(* Logix 5000 project; controller DSFW_Budzar vendor 1 type 14 code 154 rev 32.13; software revision 32.03 *)
// Unit Model Number: DSFW-0512-C-FCB-S1-SP
// Unit Serial Number: 202008-38944-1

TASK MainTask (continuous, watchdog 500 ms) : A_MainProgram, B_Process_Control, D_Refrigeration_Control
TASK PID_Fast_Loop (periodic, rate 500 ms, priority 1, watchdog 1000 ms) : Pressure_PID, EEV_PID
TASK PID_Slow_Loop (periodic, rate 1000 ms, priority 1, watchdog 500 ms) : Main

MODULES
   Local : vendor 1 type 14 code 154 (PointIO 0, rev 32.13)
      SLOT_5 : 1734-IR2 (PointIO 5, rev 3.1, Input RPI 80 ms)
           Local:5:I.Ch0Data   // TE-105 Compressor Suction Temperature (404A)
           Local:5:I.Ch1Data   // TE-204 Evaporator Suction Line Temperature
      SLOT_4 : 1734-IR2 (PointIO 4, rev 3.1, Input RPI 80 ms)
           Local:4:I.Ch0Data   // TE-103 Liquid Line Temperature (404A)
           Local:4:I.Ch1Data   // TE-104 Evaporator Suction Temperature (404A)
      SLOT_2 : vendor 1 type 115 code 210 (PointIO 2, rev 3.1, Input RPI 80 ms)
           Local:2:I.Ch2Data   // PT-103 Compressor Discharge Pressure (449a)
           Local:2:I.Ch3Data   // PT-104 Evaporator Suction Line Pressure (449a)
           Local:2:I.Ch6Data   // PT-202 Evaporator Suction Line Pressure
           Local:2:I.Ch1Data   // PT-102 Compressor Suction Pressure (449a)
           Local:2:I.Ch0Data   // PT-101 Reactor Supply Pressure
           Local:2:I.Ch4Data   // PT-105 Nitrogen/Air Pressure
           Local:2:I.Ch7Data   // TT-*** Vessel Temperature
           Local:2:I.Ch5Data   // PT-201 Condenser Loop Supply Pressure
      SLOT_6 : 1734-IR2 (PointIO 6, rev 3.1, Input RPI 80 ms)
           Local:6:I.Ch0Data   // Spare
           Local:6:I.Ch1Data   // Spare
      SLOT_3 : 1734-IR2 (PointIO 3, rev 3.1, Input RPI 80 ms)
           Local:3:I.Ch0Data   // TE-101 Reactor Supply Temperature
           Local:3:I.Ch1Data   // TE-102 Reactor Return Temperature
      SLOT_9 : 1734-IE2C (PointIO 9, rev 3.1, Input RPI 80 ms)
           Local:9:I.Ch0Data   // FIT-101 Flow Indicating Transmitter
      Discrete_IO : Embedded (PointIO 1, rev 32.11, Output RPI 20 ms)
           Local:1:I.Data.0   // ESTOP
           Local:1:I.Data.1   // Phase Monitor
           Local:1:I.Data.10   // Spare
           Local:1:I.Data.11   // Spare
           Local:1:I.Data.12   // Compressor Low Oil Level
           Local:1:I.Data.13   // Condenser Loop Heater High Temperature Status
           Local:1:I.Data.14   // Condenser Loop Pump Run Proof Status
           Local:1:I.Data.15   // Spare
           Local:1:I.Data.2   // Purge Panel
           Local:1:I.Data.3   // Process Pump Run-Proof Contact
           Local:1:I.Data.4   // Process Heater #1 High Temperature
           Local:1:I.Data.5   // Spare
           Local:1:I.Data.6   // Spare
           Local:1:I.Data.7   // Spare
           Local:1:I.Data.8   // Compressor Run-Proof Contact
           Local:1:I.Data.9   // Compressor Motor Protector
           Local:1:O.Data.0   // Process Pump Motor Start Contactor
           Local:1:O.Data.1   // Process Heater #1 Output Enable
           Local:1:O.Data.10   // Spare
           Local:1:O.Data.11   // Spare
           Local:1:O.Data.12   // Spare
           Local:1:O.Data.13   // Spare
           Local:1:O.Data.14   // Spare
           Local:1:O.Data.15   // Spare
           Local:1:O.Data.2   // Spare
           Local:1:O.Data.3   // Spare
           Local:1:O.Data.4   // Spare
           Local:1:O.Data.5   // Compressor Motor Contactor
           Local:1:O.Data.6   // Spare
           Local:1:O.Data.7   // Spare
           Local:1:O.Data.8   // Condenser Loop Pump Motor Relay
           Local:1:O.Data.9   // Spare
      SLOT_8 : vendor 1 type 115 code 211 (PointIO 8, rev 3.1, Output RPI 80 ms)
           Local:8:O.Ch2Data   // Spare
           Local:8:O.Ch3Data   // Spare
           Local:8:O.Ch1Data   // PCV-101 Condenser Pressure Control
           Local:8:O.Ch0Data   // TCV-102 Hot Gas Bypass Valve
      SLOT_7 : vendor 1 type 115 code 211 (PointIO 7, rev 3.1, Output RPI 80 ms)
           Local:7:O.Ch2Data   // EEV-102 Compressor #1 Desuperheat Valve
           Local:7:O.Ch3Data   // TCV-101 Hot Gas Bypass Valve
           Local:7:O.Ch1Data   // EEV-101 Evaporator Electric Expansion Valve
           Local:7:O.Ch0Data   // SCR-101 SCR Heater Control
END_MODULES

TYPE BL_Analog_Input :
STRUCT
   Scale_4mA : REAL;
   Scale_20mA : REAL;
   Offset : REAL;
   Output : REAL;
   Fault_Delay : DINT;
END_STRUCT
END_TYPE

ADD_ON_INSTRUCTION BudLib_Analog_Sensor   (* revision 1.0 *)
VAR_IN_OUT
   BL_Analog_Input : BL_Analog_Input; {required}
END_VAR
VAR_INPUT
   Raw_Data : REAL; {required}
   Sensor_Type : BOOL; {required}   // 0 = 4-20mA 1 = RTD
   Disable_High_Fault : BOOL; {required}
END_VAR
VAR_OUTPUT
   Sensor_Alarm : BOOL; {access None, required}
END_VAR
VAR_INPUT
   CLR_Alarm : BOOL; {required}
   Fault_Disable : BOOL; {required}   // Disable Fault
END_VAR
VAR
   Fault_Delay_TMR : TIMER; {access None}
END_VAR

ROUTINE Logic   (* ladder *)
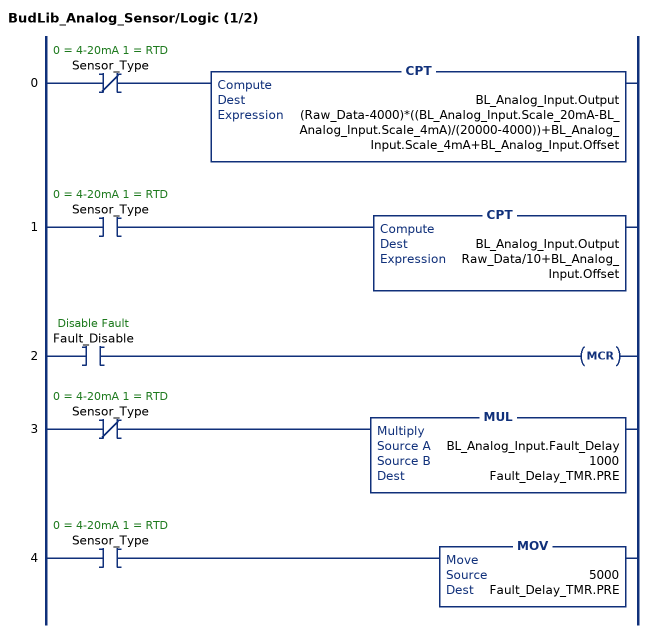
   0: XIO(Sensor_Type)CPT(BL_Analog_Input.Output,(Raw_Data-4000)*((BL_Analog_Input.Scale_20mA-BL_Analog_Input.Scale_4mA)/(20000-4000))+BL_Analog_Input.Scale_4mA+BL_Analog_Input.Offset);
   1: XIC(Sensor_Type)CPT(BL_Analog_Input.Output,Raw_Data/10+BL_Analog_Input.Offset);
   2: XIC(Fault_Disable)MCR();
   3: XIO(Sensor_Type)MUL(BL_Analog_Input.Fault_Delay,1000,Fault_Delay_TMR.PRE);
   4: XIC(Sensor_Type)MOV(5000,Fault_Delay_TMR.PRE);
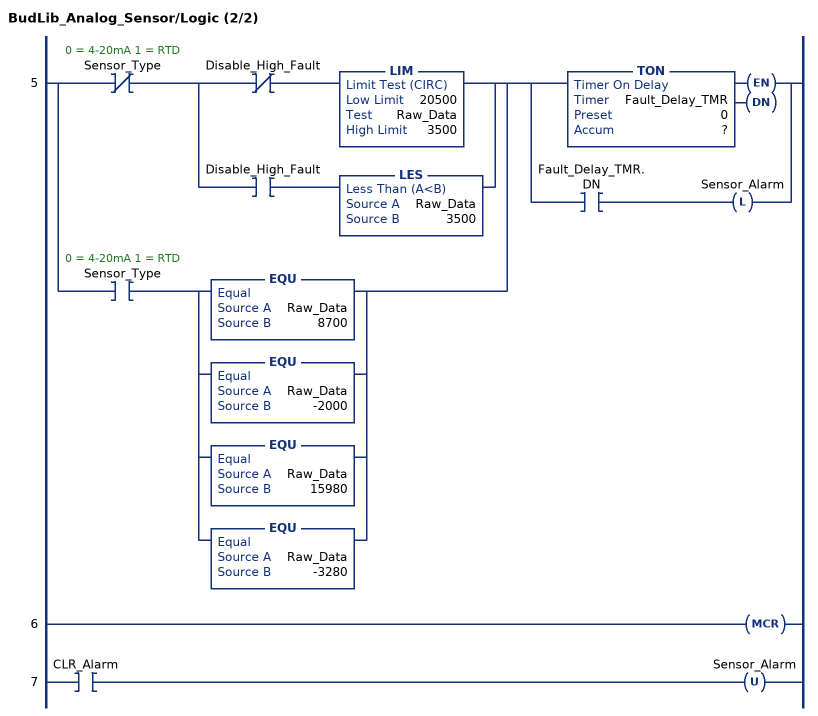
   5: [XIO(Sensor_Type) [XIO(Disable_High_Fault) LIM(20500,Raw_Data,3500) ,XIC(Disable_High_Fault) LES(Raw_Data,3500) ] ,XIC(Sensor_Type) [EQU(Raw_Data,8700) ,EQU(Raw_Data,-2000) ,EQU(Raw_Data,15980) ,EQU(Raw_Data,-3280) ] ][TON(Fault_Delay_TMR,?,?) ,XIC(Fault_Delay_TMR.DN) OTL(Sensor_Alarm) ];
   6: MCR();
   7: XIC(CLR_Alarm)OTU(Sensor_Alarm);
END_ROUTINE
END_ADD_ON_INSTRUCTION

ADD_ON_INSTRUCTION BudLib_Compressor   (* revision 1.0 *)
// Compressor Cycle and Antirecycle
VAR_OUTPUT
   PLC_Address : BOOL; {access Read Only, required}   // Compressor Start Relay
END_VAR
VAR_INPUT
   Start_Delay_Time : DINT; {required}   // Minimum Off Time, (milliseconds)
   Short_Cycle_Time : DINT; {required}   // Short Cycle Time (milliseconds)
END_VAR
VAR_OUTPUT
   Time_Remaining : DINT; {access Read Only, required}
   Compressor_Timing : BOOL; {access Read Only, required}
END_VAR
VAR_INPUT
   Compressor_OK_TO_RUN : BOOL; {access Read Only, required}
END_VAR
VAR_OUTPUT
   Start_Delay_DN : BOOL; {access Read Only}
   Start_Delay_EN : BOOL; {access Read Only}
   Start_Delay_Remaining : DINT; {access Read Only}
END_VAR
VAR
   Short_Cycle_TMR : TIMER; {access None}   // Short Cycle Timer
   Start_TMR : TIMER; {access None}   // Start Delay Timer
END_VAR

ROUTINE Logic   (* ladder *)
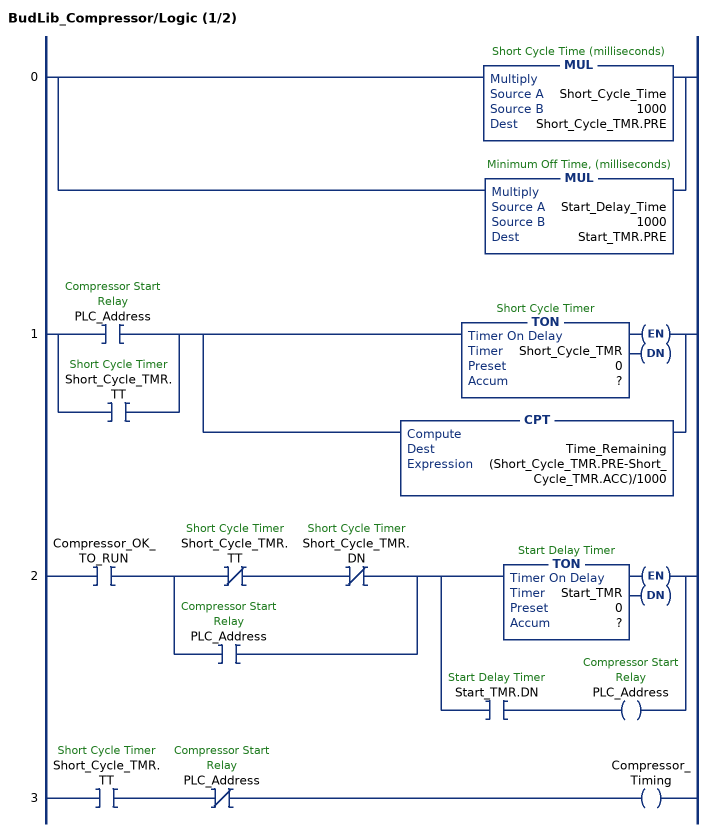
   0: [MUL(Short_Cycle_Time,1000,Short_Cycle_TMR.PRE) ,MUL(Start_Delay_Time,1000,Start_TMR.PRE) ];
   1: [XIC(PLC_Address) ,XIC(Short_Cycle_TMR.TT) ][TON(Short_Cycle_TMR,?,?) ,CPT(Time_Remaining,(Short_Cycle_TMR.PRE-Short_Cycle_TMR.ACC)/1000) ];
   2: XIC(Compressor_OK_TO_RUN)[XIO(Short_Cycle_TMR.TT) XIO(Short_Cycle_TMR.DN) ,XIC(PLC_Address) ][TON(Start_TMR,?,?) ,XIC(Start_TMR.DN) OTE(PLC_Address) ];
   3: XIC(Short_Cycle_TMR.TT)XIO(PLC_Address)OTE(Compressor_Timing);
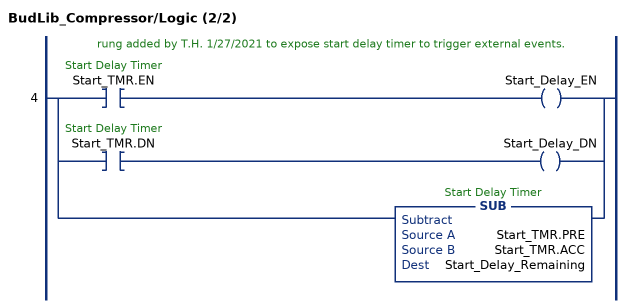
   // rung added by T.H. 1/27/2021 to expose start delay timer to trigger external events.
   4: [XIC(Start_TMR.EN) OTE(Start_Delay_EN) ,XIC(Start_TMR.DN) OTE(Start_Delay_DN) ,SUB(Start_TMR.PRE,Start_TMR.ACC,Start_Delay_Remaining) ];
END_ROUTINE
END_ADD_ON_INSTRUCTION

ADD_ON_INSTRUCTION BudLib_Heater_Step_Controller   (* revision 1.0, vendor Budzar Industries, Inc. *)
// Heaters Step Controller For Up To 10 Heaters
// Revision note:
// Initial Release 20Dec2017 (cdz)
VAR_IN_OUT
   Power_Request : REAL; {required}   // Heaters Power Request From TIC
   Heater_Circuits : DINT; {required}   // Number Of Heaters To Control (Includes SCR Controlled Heater)
   SCR : DINT; {required}   // Output To SCR scaled 0% to 100% Power
   Heater_Contactors : DINT; {required}   // Heater Contactors ON Commands (Interlock Individual Heater Circuits Outside AOI)
END_VAR
VAR_INPUT
   Interlock : BOOL; {required}   // Instruction Interlock (Sets All Outputs To Zero)
END_VAR
VAR
   Power_Total : DINT; {access None}   // Internal Calculation
   Step_Power : DINT[11]; {access None}   // Internal Calculation
END_VAR

ROUTINE Logic   (* ladder *)
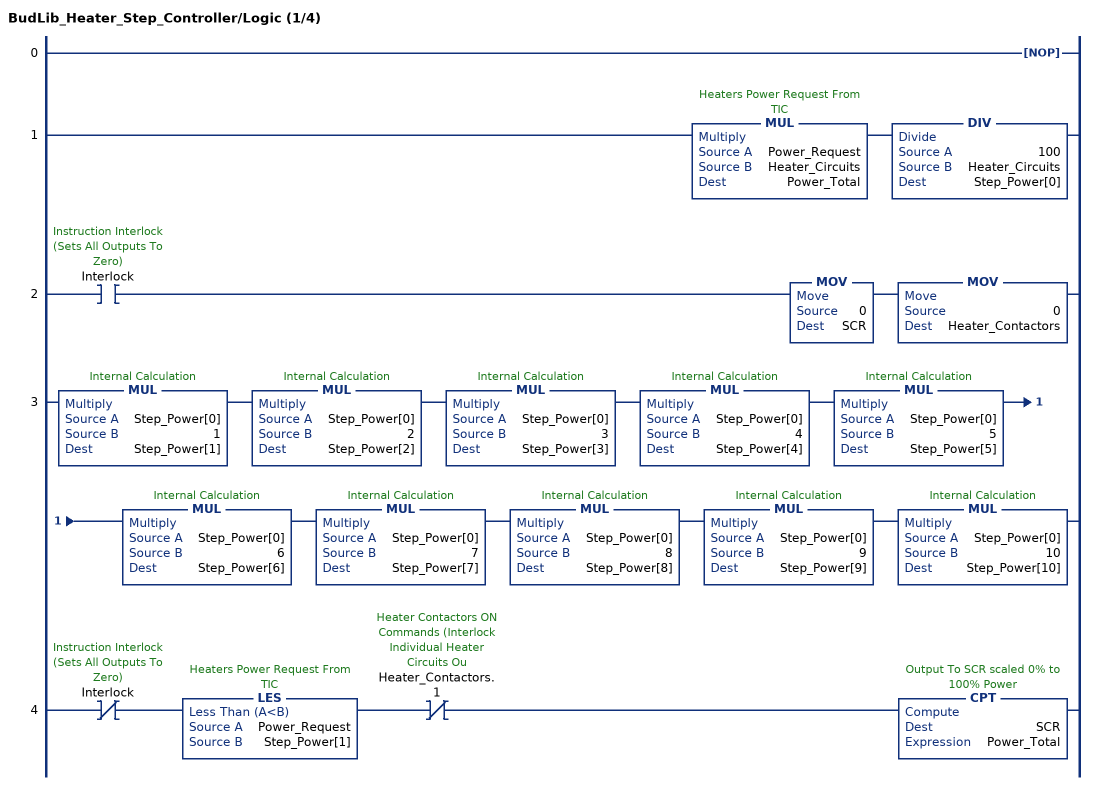
   0: NOP();
   1: MUL(Power_Request,Heater_Circuits,Power_Total)DIV(100,Heater_Circuits,Step_Power[0]);
   2: XIC(Interlock)MOV(0,SCR)MOV(0,Heater_Contactors);
   3: MUL(Step_Power[0],1,Step_Power[1])MUL(Step_Power[0],2,Step_Power[2])MUL(Step_Power[0],3,Step_Power[3])MUL(Step_Power[0],4,Step_Power[4])MUL(Step_Power[0],5,Step_Power[5])MUL(Step_Power[0],6,Step_Power[6])MUL(Step_Power[0],7,Step_Power[7])MUL(Step_Power[0],8,Step_Power[8])MUL(Step_Power[0],9,Step_Power[9])MUL(Step_Power[0],10,Step_Power[10]);
   4: XIO(Interlock)LES(Power_Request,Step_Power[1])XIO(Heater_Contactors.1)CPT(SCR,Power_Total);
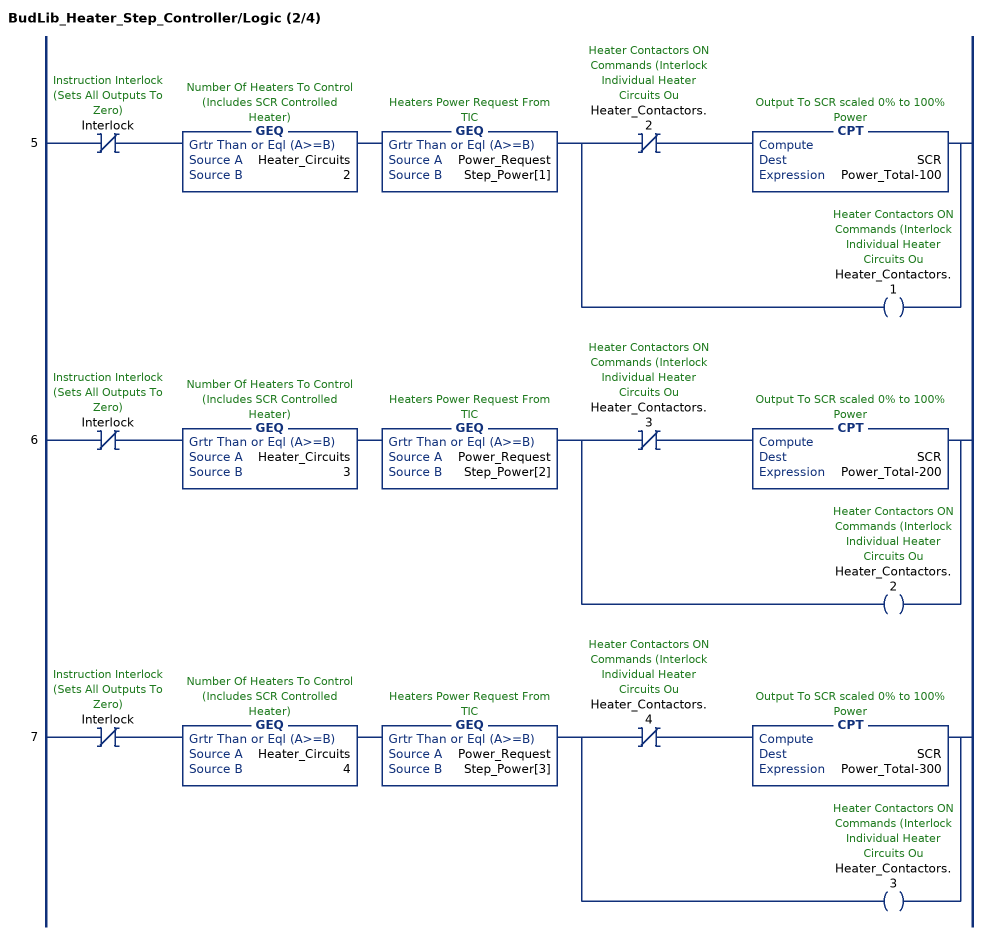
   5: XIO(Interlock)GEQ(Heater_Circuits,2)GEQ(Power_Request,Step_Power[1])[XIO(Heater_Contactors.2) CPT(SCR,Power_Total-100) ,OTE(Heater_Contactors.1) ];
   6: XIO(Interlock)GEQ(Heater_Circuits,3)GEQ(Power_Request,Step_Power[2])[XIO(Heater_Contactors.3) CPT(SCR,Power_Total-200) ,OTE(Heater_Contactors.2) ];
   7: XIO(Interlock)GEQ(Heater_Circuits,4)GEQ(Power_Request,Step_Power[3])[XIO(Heater_Contactors.4) CPT(SCR,Power_Total-300) ,OTE(Heater_Contactors.3) ];
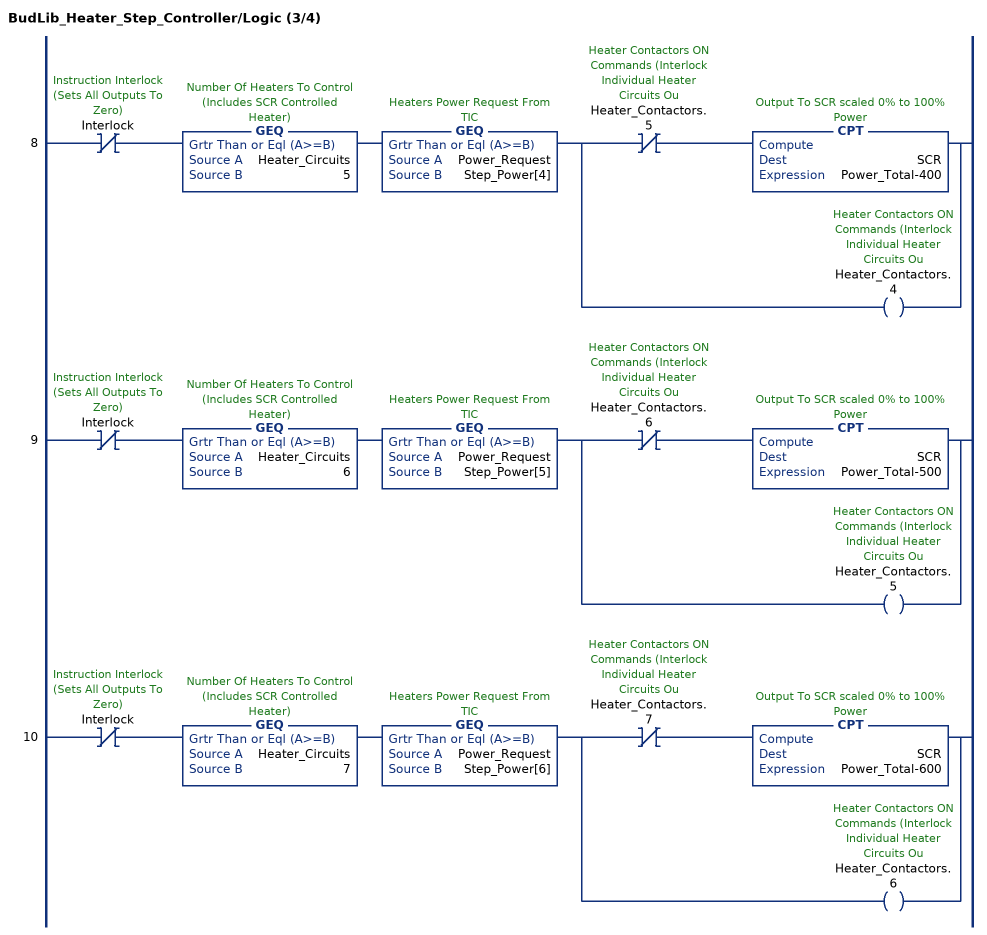
   8: XIO(Interlock)GEQ(Heater_Circuits,5)GEQ(Power_Request,Step_Power[4])[XIO(Heater_Contactors.5) CPT(SCR,Power_Total-400) ,OTE(Heater_Contactors.4) ];
   9: XIO(Interlock)GEQ(Heater_Circuits,6)GEQ(Power_Request,Step_Power[5])[XIO(Heater_Contactors.6) CPT(SCR,Power_Total-500) ,OTE(Heater_Contactors.5) ];
   10: XIO(Interlock)GEQ(Heater_Circuits,7)GEQ(Power_Request,Step_Power[6])[XIO(Heater_Contactors.7) CPT(SCR,Power_Total-600) ,OTE(Heater_Contactors.6) ];
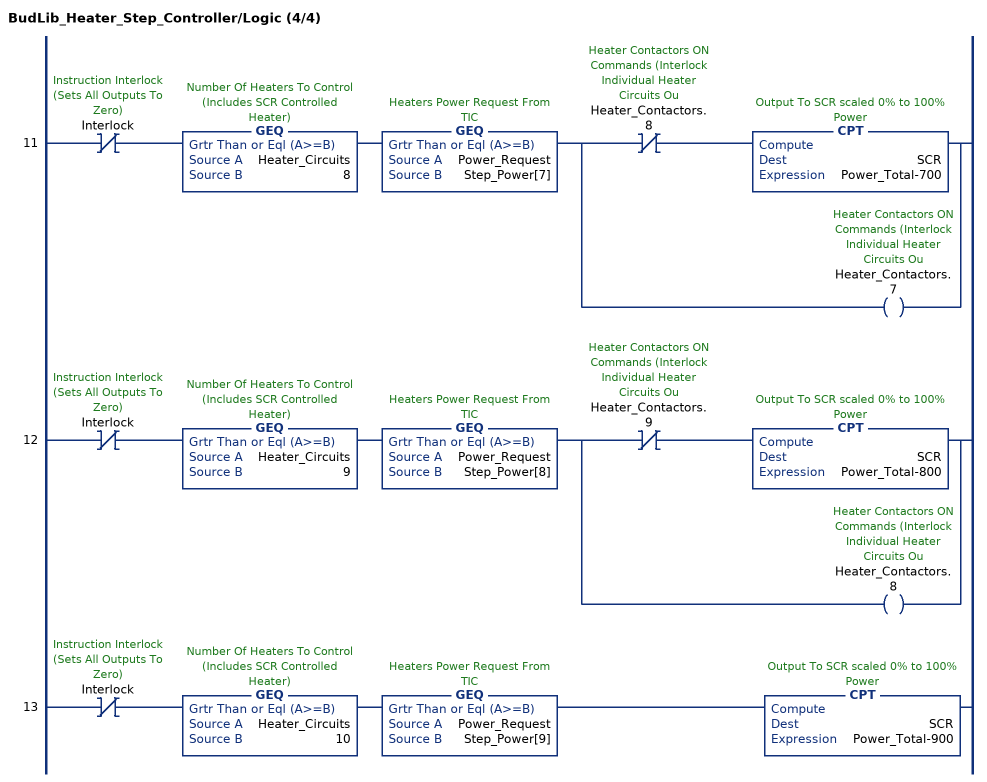
   11: XIO(Interlock)GEQ(Heater_Circuits,8)GEQ(Power_Request,Step_Power[7])[XIO(Heater_Contactors.8) CPT(SCR,Power_Total-700) ,OTE(Heater_Contactors.7) ];
   12: XIO(Interlock)GEQ(Heater_Circuits,9)GEQ(Power_Request,Step_Power[8])[XIO(Heater_Contactors.9) CPT(SCR,Power_Total-800) ,OTE(Heater_Contactors.8) ];
   13: XIO(Interlock)GEQ(Heater_Circuits,10)GEQ(Power_Request,Step_Power[9])CPT(SCR,Power_Total-900);
END_ROUTINE
END_ADD_ON_INSTRUCTION

ADD_ON_INSTRUCTION BudLib_Superheat_Subcooling   (* revision 1.2 *)
// Revision note:
// Added Refrigerant 508B
// Added Refrigerant R449A
VAR_INPUT
   Temperature : REAL; {required}   // Suction or Liquid Line Temperature
   Pressure : REAL; {required}   // Suction or Discharge Pressure
END_VAR
VAR_OUTPUT
   P2T_Suction : REAL; {access Read Only}   // Suction Pressure to Temperature Calculation
   P2T_Liquid : REAL; {access Read Only}   // Liquid Pressure to Temperature Calculation
END_VAR
VAR_INPUT
   Refridgerant_Type : INT; {required}   // 1=R-22 2=R-134a 3=R-404a 4=R-407c 5=R-407a 6=R-410a 7=R-422d 8=R-438a 9=R-507 10=R-508B 11=R-449A 12=R290
   Superheat_Subcool : BOOL; {required}   // 0 = Superheat, 1 = Subcool
END_VAR
VAR_OUTPUT
   Result : REAL; {required}   // Calculated Result
END_VAR
VAR
   Superheat : REAL; {access Read Only}   // Superheat Calculation
   Subcool : REAL; {access Read Only}   // Subcool Calculation
END_VAR

ROUTINE Logic   (* structured text *)
   
   
   Case Refridgerant_Type OF
   
   (* R-22 *)
   1:  P2T_Suction:= -0.000000165*Pressure**4 + 0.000084606*Pressure**3 - 0.016568240*Pressure**2 + 1.952262699*Pressure - 39.085397206;
       P2T_Liquid:= -0.000000165*Pressure**4 + 0.000084606*Pressure**3 - 0.016568240*Pressure**2 + 1.952262699*Pressure - 39.085397206;
   
   (*R-134a*)
   2: P2T_Suction:= -0.00000000000037678795*Pressure**6 + 0.00000000056931121499*Pressure**5 - 0.00000033878300479892*Pressure**4 + 0.00010202087796451500*Pressure**3 - 0.01710716970609380000*Pressure**2 + 1.97485706462976000*Pressure - 12.16021651744090;
      P2T_Liquid:= -0.00000000000037678795*Pressure**6 + 0.00000000056931121499*Pressure**5 - 0.00000033878300479892*Pressure**4 + 0.00010202087796451500*Pressure**3 - 0.01710716970609380000*Pressure**2 + 1.97485706462976000*Pressure - 12.16021651744090;
   
   (*R-404a*)
   3:  P2T_Suction:= -0.00000000005300893321*Pressure**6 + 0.00000002741449672112*Pressure**5 - 0.00000570303468006017*Pressure**4 + 0.00062421870492102000*Pressure**3 - 0.04148675026965520000*Pressure**2 + 2.37637660990731000000*Pressure - 49.68565233808480000000;
       P2T_Liquid:= -0.0000000000000550315164227*Pressure**6 + 0.0000000000997514242404528*Pressure**5 - 0.0000000737248710163770000*Pressure**4 + 0.0000290410699131178000000*Pressure**3- 0.0069198966935964100000000*Pressure**2  + 1.2825072984089100*Pressure - 33.916124534865200;
   
   (*R-407c*)
   4:   P2T_Suction := -0.00000000000800924737*Pressure**6 + 0.00000000557131285962*Pressure**5 - 0.00000169384905437941*Pressure**4 + 0.00028593017513500700*Pressure**3 - 0.02893370732670060000*Pressure**2 + 2.20060661934258000000*Pressure - 33.32183919094680000000;
   	P2T_Liquid:= 0.00000000000002386292*Pressure**6 - 0.00000000002645317402*Pressure**5 + 0.00000000526050718724*Pressure**4 + 0.00000470562626432580*Pressure**3 - 0.00310591635937629000*Pressure**2 + 1.00142167143801000000*Pressure - 22.25895791216770000000;
   
   (*R-407a*)
   5:	P2T_Suction:= -0.00000000011518362850*Pressure**6 + 0.00000005009100701803*Pressure**5 - 0.00000875403007261077*Pressure**4 + 0.00080807995686882400*Pressure**3 - 0.04608857801110840000*Pressure**2 + 2.36986927227190000000*Pressure - 37.26735163389090000000;
   	P2T_Liquid:= -0.00000000000003784489*Pressure**6 + 0.00000000006834533715*Pressure**5 - 0.00000005140162309636*Pressure**4 + 0.00002127640311370790*Pressure**3 - 0.00554724395898896000*Pressure**2 + 1.16486749118176000000*Pressure - 30.11932356915960000000;
   
   (*R-410a*)
   6:	P2T_Suction:= -0.00000000000007186775*Pressure**6 + 0.00000000014583668666*Pressure**5 - 0.00000011674472220023*Pressure**4 + 0.00004726707063285040*Pressure**3 - 0.01057489539488190000*Pressure**2 + 1.57409368233857000000*Pressure - 56.17353301327970000000;
   	P2T_Liquid:= -0.00000000000007186775*Pressure**6 + 0.00000000014583668666*Pressure**5 - 0.00000011674472220023*Pressure**4 + 0.00004726707063285040*Pressure**3 - 0.01057489539488190000*Pressure**2 + 1.57409368233857000000*Pressure - 56.17353301327970000000;
   
   (*R-422D*)
   7:	P2T_Suction:= 0.00000000056957976185*Pressure**5 - 0.00000058362559681170*Pressure**4 + 0.00016582335662478100*Pressure**3 - 0.02207715168838590000*Pressure**2 + 2.02610656700961000000*Pressure - 35.18819939281650000000;
   	P2T_Liquid:= 0.00000000000813454044*Pressure**5 - 0.00000001433073228086*Pressure**4 + 0.00001015786430530350*Pressure**3 - 0.00389055376093068000*Pressure**2 + 1.06625906617128000000*Pressure - 22.58790116749710000000;
   
   (*R-438a*)
   8:	P2T_Suction:= 0.00000000006078715896*Pressure**6 - 0.00000001611318229885*Pressure**5 + 0.00000020938844025320*Pressure**4 + 0.00027696642267471800*Pressure**3 - 0.03274545521389880000*Pressure**2 + 2.29322301382490000000*Pressure - 32.72178606997110000000;
   	P2T_Liquid:=  -0.00000000000003163289*Pressure**6 + 0.00000000006045751232*Pressure**5 - 0.00000004802369289111*Pressure**4 + 0.00002089758452796680*Pressure**3 - 0.00566402177639559000*Pressure**2 + 1.20642331219452000000*Pressure - 25.80440294280620000000;
   
   (*R-507*)
   9:	P2T_Suction:= -0.00000000000023273589*Pressure**6 + 0.00000000038440242299*Pressure**5 - 0.00000024966416650859*Pressure**4 + 0.00008180023458648210*Pressure**3 - 0.01483731477723890000*Pressure**2 + 1.83216631968571000000*Pressure - 49.09858575703400000000;
   	P2T_Liquid:=  -0.00000000000023273589*Pressure**6 + 0.00000000038440242299*Pressure**5 - 0.00000024966416650859*Pressure**4 + 0.00008180023458648210*Pressure**3 - 0.01483731477723890000*Pressure**2 + 1.83216631968571000000*Pressure - 49.09858575703400000000;
   
   (*R-508B*)
   10:	P2T_Suction:= -0.000000000000133667762*Pressure**6 + 0.000000000236822589*Pressure**5 - 0.000000165498946*Pressure**4 + 0.0000585053021*Pressure**3 - 0.01144174*Pressure**2 + 1.5057373*Pressure - 123.74624;
   	P2T_Liquid:=  -0.000000000000133667762*Pressure**6 + 0.000000000236822589*Pressure**5 - 0.000000165498946*Pressure**4 + 0.0000585053021*Pressure**3 - 0.01144174*Pressure**2 + 1.5057373*Pressure - 123.74624;
   
   (*R-449A*)
   11: P2T_Suction:= -0.00000000000036541159*Pressure**6 + 0.00000000054907825576*Pressure**5 - 0.00000032708993709514*Pressure**4 + 0.00009916804470212850*Pressure**3 - 0.01675694050709890000*Pressure**2 + 1.91534370751567000000*Pressure - 39.0570030049292;
   	P2T_Liquid:=  -0.00000000000036907278*Pressure**6 + 0.00000000055456970769*Pressure**5 - 0.00000033032085879095*Pressure**4 + 0.00010012437901080800*Pressure**3 - 0.01690317434666350000*Pressure**2 + 1.93545495275924000000*Pressure - 49.96916448983160000000;
   
   (*R-290*)
   12: P2T_Suction:= -8.90208426e-013*Pressure**6 + 1.11806286e-009*Pressure**5 - 5.57465512e-007*Pressure**4 + 1.42291974e-004*Pressure**3 - 0.020612964*Pressure**2 + 2.1470945*Pressure - 41.50468;
       P2T_Liquid := -8.90208426e-013*Pressure**6 + 1.11806286e-009*Pressure**5 - 5.57465512e-007*Pressure**4 + 1.42291974e-004*Pressure**3 - 0.020612964*Pressure**2 + 2.1470945*Pressure - 41.50468;
   
   END_CASE;
   
   
   IF NOT Superheat_Subcool THEN
   	Superheat:=Temperature - P2T_Suction;
   	Result := Superheat;
   
   ELSE
   	Subcool:= P2T_Liquid - Temperature;
   	Result := Subcool;
   
   END_IF;
END_ROUTINE
END_ADD_ON_INSTRUCTION

ADD_ON_INSTRUCTION P2T   (* revision 1.1 *)
// Revision note:
// Added Refrigerant 508B
VAR_INPUT
   SuctionRTD : REAL; {required}   // Suction Line RTD
   LiquidRTD : REAL; {required}   // Liquid Line RTD
   Suction_Pressure : REAL; {required}   // Compressor Suction Pressure
   Discharge_Pressure : REAL; {required}   // Compressor Discharge Pressure
END_VAR
VAR_OUTPUT
   P2T_Suction : REAL; {access Read Only}   // Suction Pressure to Temperature Calculation
   Superheat : REAL; {access Read Only, required}   // Superheat Calculation
   P2T_Liquid : REAL; {access Read Only}   // Liquid Pressure to Temperature Calculation
   Subcool : REAL; {access Read Only, required}   // Subcool Calculation
END_VAR
VAR_INPUT
   Refridgerant_Type : INT; {required}   // 1=R-22 2=R-134a 3=R-404a 4=R-407c 5=R-407a 6=R-410a 7=R-422d 8=R-438a 9=R-507 10=R-508B
END_VAR

ROUTINE Logic   (* structured text *)
   
   
   Case Refridgerant_Type OF
   
   (* R-22 *)
   1:  P2T_Suction:= -0.000000165*Suction_Pressure**4 + 0.000084606*Suction_Pressure**3 - 0.016568240*Suction_Pressure**2 + 1.952262699*Suction_Pressure - 39.085397206;
       P2T_Liquid:= -0.000000165*Discharge_Pressure**4 + 0.000084606*Discharge_Pressure**3 - 0.016568240*Discharge_Pressure**2 + 1.952262699*Discharge_Pressure - 39.085397206; ;
   
   (*R-134a*)
   2: P2T_Suction:= -0.00000000000037678795*Suction_Pressure**6 + 0.00000000056931121499*Suction_Pressure**5 - 0.00000033878300479892*Suction_Pressure**4 + 0.00010202087796451500*Suction_Pressure**3 - 0.01710716970609380000*Suction_Pressure**2 + 1.97485706462976000*Suction_Pressure - 12.16021651744090;
      P2T_Liquid:= -0.00000000000037678795*Discharge_Pressure**6 + 0.00000000056931121499*Discharge_Pressure**5 - 0.00000033878300479892*Discharge_Pressure**4 + 0.00010202087796451500*Discharge_Pressure**3 - 0.01710716970609380000*Discharge_Pressure**2 + 1.97485706462976000*Discharge_Pressure - 12.16021651744090;
   
   (*R-404a*)
   3:  P2T_Suction:= -0.00000000005300893321*Suction_Pressure**6 + 0.00000002741449672112*Suction_Pressure**5 - 0.00000570303468006017*Suction_Pressure**4 + 0.00062421870492102000*Suction_Pressure**3 - 0.04148675026965520000*Suction_Pressure**2 + 2.37637660990731000000*Suction_Pressure - 49.68565233808480000000;
       P2T_Liquid:= -0.0000000000000550315164227*Discharge_Pressure**6 + 0.0000000000997514242404528*Discharge_Pressure**5 - 0.0000000737248710163770000*Discharge_Pressure**4 + 0.0000290410699131178000000*Discharge_Pressure**3- 0.0069198966935964100000000*Discharge_Pressure**2  + 1.2825072984089100*Discharge_Pressure - 33.916124534865200;
   
   (*R-407c*)
   4:   P2T_Suction := -0.00000000000800924737*Suction_Pressure**6 + 0.00000000557131285962*Suction_Pressure**5 - 0.00000169384905437941*Suction_Pressure**4 + 0.00028593017513500700*Suction_Pressure**3 - 0.02893370732670060000*Suction_Pressure**2 + 2.20060661934258000000*Suction_Pressure - 33.32183919094680000000;
   	P2T_Liquid:= 0.00000000000002386292*Discharge_Pressure**6 - 0.00000000002645317402*Discharge_Pressure**5 + 0.00000000526050718724*Discharge_Pressure**4 + 0.00000470562626432580*Discharge_Pressure**3 - 0.00310591635937629000*Discharge_Pressure**2 + 1.00142167143801000000*Discharge_Pressure - 22.25895791216770000000;
   
   (*R-407a*)
   5:	P2T_Suction:= -0.00000000011518362850*Suction_Pressure**6 + 0.00000005009100701803*Suction_Pressure**5 - 0.00000875403007261077*Suction_Pressure**4 + 0.00080807995686882400*Suction_Pressure**3 - 0.04608857801110840000*Suction_Pressure**2 + 2.36986927227190000000*Suction_Pressure - 37.26735163389090000000;
   	P2T_Liquid:= -0.00000000000003784489*Discharge_Pressure**6 + 0.00000000006834533715*Discharge_Pressure**5 - 0.00000005140162309636*Discharge_Pressure**4 + 0.00002127640311370790*Discharge_Pressure**3 - 0.00554724395898896000*Discharge_Pressure**2 + 1.16486749118176000000*Discharge_Pressure - 30.11932356915960000000;
   
   (*R-410a*)
   6:	P2T_Suction:= -0.00000000000007186775*Suction_Pressure**6 + 0.00000000014583668666*Suction_Pressure**5 - 0.00000011674472220023*Suction_Pressure**4 + 0.00004726707063285040*Suction_Pressure**3 - 0.01057489539488190000*Suction_Pressure**2 + 1.57409368233857000000*Suction_Pressure - 56.17353301327970000000;
   	P2T_Liquid:= -0.00000000000007186775*Discharge_Pressure**6 + 0.00000000014583668666*Discharge_Pressure**5 - 0.00000011674472220023*Discharge_Pressure**4 + 0.00004726707063285040*Discharge_Pressure**3 - 0.01057489539488190000*Discharge_Pressure**2 + 1.57409368233857000000*Discharge_Pressure - 56.17353301327970000000;
   
   (*R-422D*)
   7:	P2T_Suction:= 0.00000000056957976185*Suction_Pressure**5 - 0.00000058362559681170*Suction_Pressure**4 + 0.00016582335662478100*Suction_Pressure**3 - 0.02207715168838590000*Suction_Pressure**2 + 2.02610656700961000000*Suction_Pressure - 35.18819939281650000000;
   	P2T_Liquid:= 0.00000000000813454044*Discharge_Pressure**5 - 0.00000001433073228086*Discharge_Pressure**4 + 0.00001015786430530350*Discharge_Pressure**3 - 0.00389055376093068000*Discharge_Pressure**2 + 1.06625906617128000000*Discharge_Pressure - 22.58790116749710000000;
   
   (*R-438a*)
   8:	P2T_Suction:= 0.00000000006078715896*Suction_Pressure**6 - 0.00000001611318229885*Suction_Pressure**5 + 0.00000020938844025320*Suction_Pressure**4 + 0.00027696642267471800*Suction_Pressure**3 - 0.03274545521389880000*Suction_Pressure**2 + 2.29322301382490000000*Suction_Pressure - 32.72178606997110000000;
   	P2T_Liquid:=  -0.00000000000003163289*Discharge_Pressure**6 + 0.00000000006045751232*Discharge_Pressure**5 - 0.00000004802369289111*Discharge_Pressure**4 + 0.00002089758452796680*Discharge_Pressure**3 - 0.00566402177639559000*Discharge_Pressure**2 + 1.20642331219452000000*Discharge_Pressure - 25.80440294280620000000;
   
   (*R-507*)
   9:	P2T_Suction:= -0.00000000000023273589*Suction_Pressure**6 + 0.00000000038440242299*Suction_Pressure**5 - 0.00000024966416650859*Suction_Pressure**4 + 0.00008180023458648210*Suction_Pressure**3 - 0.01483731477723890000*Suction_Pressure**2 + 1.83216631968571000000*Suction_Pressure - 49.09858575703400000000;
   	P2T_Liquid:=  -0.00000000000023273589*Discharge_Pressure**6 + 0.00000000038440242299*Discharge_Pressure**5 - 0.00000024966416650859*Discharge_Pressure**4 + 0.00008180023458648210*Discharge_Pressure**3 - 0.01483731477723890000*Discharge_Pressure**2 + 1.83216631968571000000*Discharge_Pressure - 49.09858575703400000000;
   
   (*R-508B*)
   10:	P2T_Suction:= -0.000000000000133667762*Suction_Pressure**6 + 0.000000000236822589*Suction_Pressure**5 - 0.000000165498946*Suction_Pressure**4 + 0.0000585053021*Suction_Pressure**3 - 0.01144174*Suction_Pressure**2 + 1.5057373*Suction_Pressure - 123.74624;
   	P2T_Liquid:=  -0.000000000000133667762*Discharge_Pressure**6 + 0.000000000236822589*Discharge_Pressure**5 - 0.000000165498946*Discharge_Pressure**4 + 0.0000585053021*Discharge_Pressure**3 - 0.01144174*Discharge_Pressure**2 + 1.5057373*Discharge_Pressure - 123.74624;
   
   
   END_CASE;
   
   Superheat:=SuctionRTD - P2T_Suction;
   
   Subcool:= P2T_Liquid - LiquidRTD;
   
END_ROUTINE
END_ADD_ON_INSTRUCTION

VAR_GLOBAL   (* controller tags *)
   ACKNOWLEDGE_ALARMS : BOOL;
   Active_Setpoint : REAL := 20.0;
   ALARMS : DINT[5] := ([1] := 2#0000_0001_0000_0000_0000_0000_0000_0000);
        [0]   // SENSOR ALARMS
        [0].0   // PT-101 Process Supply Pressure Sensor Fault
        [0].1   // PT-102 404A Compressor Suction Pressure Sensor Fault
        [0].10   // TE-101 Process Supply Temperature Sensor Fault
        [0].11   // TE-102 Process Return Temperature Sensor Fault
        [0].12   // TE-103 404A Liquid Line Temperature Sensor Fault
        [0].13   // TE-104 404A Evaporator Suction Temperature Sensor Fault
        [0].14   // TE-105 404A Compressor Suction Temperature Sensor Fault
        [0].15   // TE-106 Condenser Chilled Water Outlet Temperature Sensor Fault
        [0].16   // TE-108 Condenser Chilled Water Inlet Temperature Sensor Fault
        [0].2   // PT-103 404A Compressor Discharge Pressure Sensor Fault
        [0].3   // PT-104 404A Evaporator Suction Line Pressure Sensor Fault
        [0].4   // PT-105 4 MTR-101 Low Suction Pressure Sensor Fault
        [0].5   // FIT-101 Process Supply Flow Transmitter Fault
        [0].6   // PT-107 Pump Suction Pressure Sensor Fault
        [0].7   // PT-108 Pump Discharge Pressure Sensor Fault
        [0].9   // TT-*** Vessel Temperature Transmitter Sensor Fault
        [1]   // General/Process Alarms
        [1].0   // Process Pump Run-Proof Alarm
        [1].1   // Heater #1 Elements High Temperature Alarm
        [1].10   // Jacket High High Temperature Alarm
        [1].11   // Jacket HighTemperature Alarm
        [1].12   // Vessel Low Low Temperature Alarm
        [1].13   // Spare
        [1].14   // Vessel High High Temperature Alarm
        [1].15   // Jacket/Vessel High Delta T Alarm
        [1].16   // Glycol Tank Low Level Alarm
        [1].17   // Process Pump Low Suction Pressure Alarm
        [1].18   // Spare
        [1].19   // Spare
        [1].2   // Spare
        [1].20   // Purge Panel Low Pressure
        [1].21   // Spare
        [1].23   // Remote Temperature Setpoint from Plant DCS is out-of-range
        [1].24   // DCS Communication Fault
        [1].25   // Condenser Water Inlet Temperature High Alarm
        [1].3   // Phase Monitor Fault
        [1].4   // Emergency Stop
        [1].5   // Process Pump Low Pressure Alarm
        [1].6   // Process Pump High Pressure Alarm
        [1].8   // Jacket Low Low Temperature Alarm
        [1].9   // Jacket Low Temperature Alarm
        [2]   // R404A Refrigeration Alarms
        [2].0   // Compressor Run-Proof Alarm
        [2].1   // Compressor Low Pressure
        [2].11   // PT-202 CONDENSER EVAPORATOR SUCTION LINE PRESSURE TRANSMITTER ALARM
        [2].12   // TE-201 CONDENSER LOOP SUPPLY TEMPERATURE SENSOR FAULT
        [2].13   // TE-202 CONDENSER LOOP RETURN TEMPERATURE SENSOR FAULT
        [2].14   // TE-204 EVAPORATOR SUCTION LINE TEMPERATURE SENSOR FAULT
        [2].2   // Compressor High Pressure
        [2].3   // Low Superheat
        [2].4   // High Superheat
        [2].5   // Compressor Low Oil Level
        [2].6   // Compressor Motor Protector
        [2].7   // Condening Glycol/Water Temmperature Too High Alarm
        [4]   // Module Faults
        [4].0   // PLC101 SLOT 2 1734-IE8C MODULE CRASH
        [4].1   // PLC101 SLOT 3 1734-IR2 MODULE CRASH
        [4].2   // PLC101 SLOT 4 1734-IR2 MODULE CRASH
        [4].3   // PLC101 SLOT 5 1734-IR2 MODULE CRASH
        [4].4   // PLC101 SLOT 6 1734-IR2 MODULE CRASH
        [4].5   // PLC101 SLOT 7 1734-OE4C MODULE CRASH
        [4].6   // PLC101 SLOT 8 1734-OE4C MODULE CRASH
        [4].7   // PLC101 SLOT 9 1734-IE2C MODULE CRASH
   ALARMS_PRESENT : BOOL := 1;
   ALWAYS_OFF : BOOL;
   Batch_High_High_Temp_Delay : TIMER := (PRE := 30000);
   Batch_High_High_Temp_Setpoint : REAL;
   Batch_High_Temp_Setpoint : REAL;
   Batch_Jacket_DT_Temp_Delay : TIMER := (PRE := 30000);
   Batch_Low_Low_Temp_Delay : TIMER := (PRE := 30000);
   Batch_Low_Low_Temp_Setpoint : REAL := -10.0;
   Batch_Low_Temp_Delay : TIMER := (PRE := 5000);
   Batch_Low_Temp_Setpoint : REAL;
   Batch_Mode_Enable : BOOL;
   Batch_Mode_Running : BOOL;
   Blanket_Pressure_Delta_PV : REAL := 0.95624924;
   BudLib_P2T_1 : BudLib_Superheat_Subcooling := (Temperature := 85.1, Pressure := 110.7004, P2T_Suction := 53.529312, P2T_Liquid := 53.13972, Refridgerant_Type := 3, Result := 31.570686);
   BudLib_P2T_2 : BudLib_Superheat_Subcooling := (Temperature := 73.7, Pressure := 163.45125, P2T_Suction := 73.087265, P2T_Liquid := 75.620316, Refridgerant_Type := 3, Superheat_Subcool := 1, Result := 1.9203186);
   BudLib_P2T_3 : BudLib_Superheat_Subcooling := (Temperature := 75.1, Pressure := 110.693596, P2T_Suction := 53.524734, P2T_Liquid := 53.136364, Refridgerant_Type := 3, Result := 21.575264);
   BudLib_P2T_4 : BudLib_Superheat_Subcooling := (Temperature := 26.4, Pressure := 24.42431, P2T_Suction := -9.100571, P2T_Liquid := -6.3220596, Refridgerant_Type := 3, Result := 35.500572);
   C1_Low_Oil_Timer : TIMER := (PRE := 5000);
   C1_MP_Timer : TIMER := (PRE := 3000);
   C1_Run_Proof_Timer : TIMER := (PRE := 3000);
   C2_MP_Timer : TIMER := (PRE := 3000);
   C2_Run_Proof_Timer : TIMER := (PRE := 3000);
   C3_MP_Timer : TIMER := (PRE := 3000);
   C3_Run_Proof_Timer : TIMER := (PRE := 3000);
   C_101_AUX : ALIAS FOR Local:1:I.Data.8;
   CLR_Alarms : BOOL;
   Comp_1 : BudLib_Compressor := (Start_Delay_Time := 10, Short_Cycle_Time := 300, Start_Delay_Remaining := 10000);   // R507A Compressor 1
   Comp_1_Status : BOOL;
   Comp_404A_Timing_1 : BOOL;
   Comp_404A_Timing_2 : BOOL;
   Comp_Start_Purge_Relay : BOOL;
   Compressor_R404A_Subcooling : REAL := 1.9203186;
   Compressor_R404A_Superheat : REAL := 31.570686;
   Compressor_Start_Request : BOOL;
   Condenser_Water_Inlet_Temp_Limit : REAL := 100.0;
   Condenser_Water_Inlet_Temp_TMR : TIMER := (PRE := 10000);
   CR_002 : ALIAS FOR Local:1:I.Data.0;   // Emergency Stop Safety Relay Status
   CR_003 : ALIAS FOR Local:1:O.Data.15;   // General Fault Relay
   CR_01 : ALIAS FOR Local:1:I.Data.15;   // Glycol Tank Low Level Alarm Relay Dry Contact
   CR_108 : ALIAS FOR Local:1:O.Data.0;   // Process Pump Motor Relay (Energizes Contactor M-101)
   CR_109 : ALIAS FOR Local:1:O.Data.5;   // Compressor Motor Relay (Energizes Contactor C-101)
   CR_201 : ALIAS FOR Local:1:O.Data.8;   // GFS-10 Auto Start Relay (Enables Glycol Pump)
   DCS_Comm_TMR : TIMER := (PRE := 10000, ACC := 10000, EN := 1, DN := 1);
   DCS_Heartbeat_Returned : DINT;
   DCS_Heartbeat_Returned_Last : DINT;
   EEV_101_Auto_Manual : BOOL;
   EEV_101_High_Range_CV_Max : REAL := 65.0;
   EEV_101_High_Range_CV_Min : REAL := 9.0;
   EEV_101_Low_Range_CV_Max : REAL := 88.0;
   EEV_101_Low_Range_CV_Min : REAL := 5.0;
   EEV_101_Manual_Percent : REAL := 100.0;
   EEV_101_Mid_Range_CV_Max : REAL := 87.0;
   EEV_101_Mid_Range_CV_Min : REAL := 8.0;
   EEV_101_Pressure_PIDE : PID_ENHANCED := (PV := 110.693596, PVEUMax := 121.5, PVEUMin := -27.3, SPProg := 100.0, SPOper := 100.0, SPHLimit := 121.5, SPLLimit := -27.3, RatioProg := 1.0, RatioOper := 1.0, RatioHLimit := 1.0, RatioLLimit := 1.0, CVEUMax := 20000.0, CVEUMin := 4000.0, CVHLimit := 87.0, CVLLimit := 8.0, HandFB := 100.0, PGain := 3.0, IGain := 8.0, PVEDerivative := 1, ProgOverrideReq := 1, RTSTime := 1, CVEU := 4000.0, CVLAlarm := 1, SP := 100.0, SPPercent := 85.55108, PVPercent := 92.737625, E := -10.693596, EPercent := -7.1865463, InitPrimary := 1, WindupLOut := 1, Ratio := 1.0, ProgOper := 1, Override := 1, DeltaT := 0.5);
   EEV_101_Pressure_Setpoint : REAL := 100.0;
   EEV_101_Run_PIDE : BOOL;
   EEV_101_Run_Temp_PIDE : BOOL;
   EEV_101_SH_PIDE : PID_ENHANCED := (PV := 21.575264, PVEUMax := 200.0, PVEUMin := -100.0, SPProg := 12.0, SPOper := 12.0, SPHLimit := 200.0, SPLLimit := -100.0, RatioProg := 1.0, RatioOper := 1.0, RatioHLimit := 1.0, RatioLLimit := 1.0, CVEUMax := 20000.0, CVEUMin := 4000.0, CVHLimit := 87.0, CVLLimit := 8.0, HandFB := 100.0, ControlAction := 1, PGain := 5.0, IGain := 12.0, PVEDerivative := 1, ProgOverrideReq := 1, RTSTime := 1, CVEU := 4000.0, CVLAlarm := 1, SP := 12.0, SPPercent := 37.333332, PVPercent := 40.52509, E := 9.575264, EPercent := 3.1917572, InitPrimary := 1, WindupHOut := 1, Ratio := 1.0, ProgOper := 1, Override := 1, DeltaT := 0.5);
   EEV_101_Stop_PIDE : BOOL := 1;
   EEV_101_Superheat_Setpoint : REAL := 12.0;
   EEV_101_Temperature_PIDE : PID_ENHANCED := (PV := 23.3, PVEUMax := 200.0, PVEUMin := -40.0, SPProg := 20.0, SPOper := 23.3, SPCascade := 23.3, SPHLimit := 200.0, SPLLimit := -40.0, RatioProg := 1.0, RatioOper := 1.0, RatioHLimit := 1.0, RatioLLimit := 1.0, CVEUMax := 20000.0, CVEUMin := 4000.0, CVHLimit := 87.0, CVLLimit := 8.0, HandFB := 100.0, ControlAction := 1, PGain := 3.0, IGain := 8.0, PVEDerivative := 1, PVTracking := 1, AllowCasRat := 1, ProgOverrideReq := 1, RTSTime := 1, CVEU := 4000.0, CVLAlarm := 1, SP := 23.3, SPPercent := 26.374998, PVPercent := 26.374998, InitPrimary := 1, WindupHOut := 1, Ratio := 1.0, ProgOper := 1, Override := 1, DeltaT := 0.5);
   EEV_101_To_Purge : BOOL;   // Oil Management, Call For Purge with EEV-101
   EEV_102_Auto_Manual : BOOL;
   EEV_102_Manual_Percent : REAL;
   EEV_102_PIDE : PID_ENHANCED := (PV := 31.570686, PVEUMax := 200.0, PVEUMin := -40.0, SPProg := 40.0, SPOper := 31.570686, SPHLimit := 200.0, SPLLimit := -40.0, RatioProg := 1.0, RatioOper := 1.0, RatioHLimit := 1.0, RatioLLimit := 1.0, CVEUMax := 20000.0, CVEUMin := 4000.0, CVHLimit := 100.0, ControlAction := 1, PGain := 2.0, IGain := 3.0, PVEDerivative := 1, PVTracking := 1, ProgOverrideReq := 1, RTSTime := 1, CVEU := 4000.0, SP := 31.570686, SPPercent := 29.82112, PVPercent := 29.82112, InitPrimary := 1, Ratio := 1.0, ProgOper := 1, Override := 1, DeltaT := 0.5);
   EEV_102_Run_PIDE : BOOL;
   EEV_102_Stop_PIDE : BOOL := 1;
   EEV_102_Superheat_Setpoint : REAL := 40.0;
   EEV_201_Auto_Manual : BOOL;
   EEV_High_Range_Max_Temp : REAL := 90.0;
   EEV_High_Range_Min_Temp : REAL := 55.1;
   EEV_Low_Range_Max_Temp : REAL := -5.0;
   EEV_Low_Range_Min_Temp : REAL := -10.0;
   EEV_Manual_Relief_Delay : TIMER := (PRE := 75000);   // Oil Management, Delay until Flush begins
   EEV_Manual_Relief_Timer : TIMER := (PRE := 15000);   // Oil Management, Duration of Flush
   EEV_Mid_Range_Max_Temp : REAL := 55.0;
   EEV_Mid_Range_Min_Temp : REAL := -4.1;
   Enable_Batch : BOOL;   // Batch/Jacket Mode 0=Jacket 1=Batch
   Engineering_Alarm_Reset : TIMER := (PRE := 10000);
   Evaporator_R404A_Superheat : REAL := 21.575264;
   F8 : REAL[48] := ([0] := 24.885624, [2] := 0.033749998, [3] := 22.1, [5] := 23.3, [6] := 25.1575, [7] := 24.813124, [8] := 110.693596, [9] := 75.1, [10] := 85.1, [11] := 110.7004, [12] := 73.7, [13] := 163.45125, [14] := 73.4, [15] := 28.827812, [16] := 71.5, [17] := 47.85, [23] := 20.0, [28] := 25.0); {produced}   // FLOAT DATA FOR PLANT SUPERVISORY SYSTEM
   FCV_101 : ALIAS FOR Local:8:O.Ch2Data;   // Process Bypass Flow Control Valve
   FIC_101_Manual_Percent : REAL := 50.0;
   FIC_101_PIDE : PID_ENHANCED := (PV := 0.031875, PVEUMax := 165.0, PVEUMin := -20.0, SPProg := 20.0, SPOper := 0.031875, SPHLimit := 165.0, SPLLimit := -20.0, RatioProg := 1.0, RatioOper := 1.0, RatioHLimit := 1.0, RatioLLimit := 1.0, CVEUMax := 20000.0, CVEUMin := 4000.0, CVHLimit := 100.0, HandFB := 50.0, PGain := 1.2, IGain := 25.0, PVEDerivative := 1, PVTracking := 1, ProgOverrideReq := 1, RTSTime := 1, CVEU := 4000.0, SP := 0.031875, SPPercent := 10.82804, PVPercent := 10.82804, InitPrimary := 1, Ratio := 1.0, ProgOper := 1, Override := 1, DeltaT := 0.5);
   FIC_101_Run_PID : BOOL;
   FIC_101_Setpoint : REAL := 20.0;
   FIC_101_Stop_PID : BOOL := 1;
   FIT_101 : BL_Analog_Input := (Scale_20mA := 30.0, Output := 0.031875);   // Flow Indicating Transmitter
   FIT_101_PID_Scale_Max : REAL := 165.0;
   FIT_101_PID_Scale_Min : REAL := -20.0;
   Glycol_Pump_Disable_TMR : TIMER := (PRE := 10000);   // Disable Glycol Fill Pump on High PSI (backup for Pressure Switch on Neptune)
   Heater_Contactors : DINT;
   Heater_Step_Controller : BudLib_Heater_Step_Controller := (Interlock := 1);
   High_Range_Max_Temp : REAL := 90.0;
   High_Range_Min_Temp : REAL := 55.1;
   HMI_Batch_Hi_Hi_Temp_Delay : DINT := 30;
   HMI_Batch_Jacket_DT_Temp_Delay : DINT := 30;
   HMI_Batch_Low_Low_Temp_Delay : DINT := 30;
   HMI_Bypass_Speed : DINT := 3;
   HMI_Bypass_Status : BOOL;
   HMI_Condenser_Water_Inlet_Temp_Delay : DINT := 10;
   HMI_EEV_101_CV : REAL;
   HMI_EEV_101_Lamp : BOOL;
   HMI_EEV_102_CV : REAL;
   HMI_EEV_102_Lamp : BOOL;
   HMI_EEV_Manual_Relief_Delay : REAL := 75.0;   // Oil Management, Delay to start relief entered in minutes.
   HMI_EEV_Manual_Relief_Timer : REAL := 15.0;   // Oil Management, Relief Duration entered in seconds
   HMI_FCV_101_CV : REAL;
   HMI_FCV_101_Lamp : BOOL;
   HMI_Heater_1_Lamp : BOOL;
   HMI_Heater_2_Lamp : BOOL;
   HMI_Jacket_Hi_Hi_Temp_Delay : DINT := 30;
   HMI_Jacket_Hi_Temp_Delay : REAL := 30.0;
   HMI_Jacket_Low_Low_Temp_Delay : DINT := 30;
   HMI_Jacket_Low_Temp_Delay : REAL := 30.0;
   HMI_Low_Pump_Suction_Pressure_Delay : REAL := 30.0;
   HMI_Low_Suction_Pressure_Delay : DINT := 10;
   HMI_Oil_Purge_Retries_Reset_Min : REAL := 10.0;   // Oil Management, Compressor Runtime before resetting retry accumulator
   HMI_PCV_101_Flush_Time : DINT := 30;
   HMI_PCV_101_Lamp : BOOL;
   HMI_PCV_101_Output : REAL;
   HMI_Pump_Start : BOOL;
   HMI_Pump_Status : BOOL;
   HMI_Pump_Stop : BOOL;
   HMI_R404A_Hot_Gas_Switch_Delay : REAL := 10.0;
   HMI_R404A_TCV_Toggle_SP : REAL := 60.0;
   HMI_R404A_Valve_Flush_SP : REAL := 80.0;   // Oil Management, desired valve position for Flush (0-100%)
   HMI_R507A_High_Superheat_Timer : DINT := 120;
   HMI_R507A_Low_Pressure_Delay : DINT := 120;
   HMI_R507A_Low_Superheat_Timer : DINT := 120;
   HMI_Ramping : BOOL;
   HMI_Remote_State_1 : BOOL;
   HMI_Remote_State_2 : BOOL;
   HMI_Return_Trend_Limits : REAL[2] := ([0] := -7.8999996, [1] := 52.1);
   HMI_SCR_Max : DINT;
   HMI_Soaking : BOOL;
   HMI_SP_Trend_Limits : REAL[2] := ([0] := -10.0, [1] := 50.0);
   HMI_Supply_Flow_Speed : DINT := 3;
   HMI_Supply_Flow_Status : BOOL;
   HMI_Supply_Trend_Limits : REAL[2] := ([0] := -6.700001, [1] := 53.3);
   HMI_TCV_101_CV : REAL;
   HMI_TCV_101_Lamp : BOOL;
   HMI_TCV_102_CV : REAL;
   HMI_TCV_102_Lamp : BOOL;
   HMI_TCV_Manual_Relief_Delay : REAL := 60.0;
   HMI_TCV_Manual_Relief_Timer : REAL := 10.0;
   HMI_Trend_Data : REAL[3] := ([0] := 20.0, [1] := 23.3, [2] := 22.1);
        [0]   // Temperature Setpoint
        [1]   // Process Supply Temperature
        [2]   // Process Return Temperature
   HMI_Valve_Flush_SP : REAL := 60.0;
   Jacket_Batch_Delta_T : REAL := 132.44063;
   Jacket_Batch_High_Delta_T_Setpoint : REAL := 100.0;
   Jacket_High_High_Temp_Delay : TIMER := (PRE := 30000);
   Jacket_High_High_Temp_Setpoint : REAL := 100.0;
   Jacket_High_Temp_Delay : TIMER := (PRE := 30000);
   Jacket_High_Temp_Setpoint : REAL := 90.0;
   Jacket_Low_Low_Temp_Delay : TIMER := (PRE := 30000);
   Jacket_Low_Low_Temp_Setpoint : REAL := -20.0;
   Jacket_Low_Temp_Delay : TIMER := (PRE := 30000);
   Jacket_Low_Temp_Setpoint : REAL := -10.0;
   Local_System_Start : BOOL;   // Local System Start 0=Stop 1=Start
   Local_Temp_Setpoint : REAL := 20.0;   // Local Temperature Setpoint
   Low_Pump_Suction_Pressure_Delay : TIMER := (PRE := 30000);
   Low_Pump_Suction_Pressure_Setpoint : REAL := 4.0;
   Low_Range_Max_Temp : REAL;
   Low_Range_Min_Temp : REAL := -10.0;
   M_101_AUX : ALIAS FOR Local:1:I.Data.3;
   Mid_Range_Max_Temp : REAL := 55.0;
   Mid_Range_Min_Temp : REAL := 0.1;
   N7 : INT[16] := ([0] := 26, [1] := 32, [10] := 60, [11] := 2); {produced}   // INTEGER DATA FOR PLANT SUPERVISORY SYSTEM
        [11].0   // REMOTE START PUSH BUTTON
        [11].1   // REMOTE STOP PUSH BUTTON
   New_Alarm_TMR : TIMER := (PRE := 500);
   NEW_ALARMS : DINT[5];   // New Alarms this scan
   NEW_ALARMS_PRESENT : BOOL;   // New Alarm Present This Scan
   NOT_ALARMS_LAST : DINT[5] := ([0] := -1, [1] := -16777217, [2] := -1, [3] := -1, [4] := -1);   // Logical NOT of Alarms Last Scan
   Num_Heaters : DINT := 2;
   Oil_Purge_Fail : BOOL;   // Oil Management, This coil will energize after configured purge retries fail
   Oil_Purge_Relay : BOOL;   // Oil Management, Oil Purge Sequence Latch
   Oil_Purge_Retires_Enable : BOOL;
   Oil_Purge_Retries_ACC : DINT;   // Oil Management, Accumulated Oil Purges this low level
   Oil_Purge_Retries_Reset : TIMER := (PRE := 600000);   // Oil Management, Reset Accumulator with 10-min without Low Level
   Oil_Purge_Retries_Reset1 : TIMER := (PRE := 10000, ACC := 10002, EN := 1, DN := 1);   // Oil Management, Used to reset accuulated retries if compressor off.
   Oil_Purge_Retries_Reset_Remaining : REAL;   // Oil Management, Time remaining until reset retries accum
   Oil_Purge_Retries_SP : DINT := 6;   // Oil Management, Desired Oil Purge Retries before Fault
   OMB_101 : ALIAS FOR Local:1:I.Data.12;
   ONS : DINT[3] := ([0] := 5);   // One-Shots
   P2T_507A : P2T := (SuctionRTD := 66.4, LiquidRTD := 61.8, Suction_Pressure := 76.8296, Discharge_Pressure := 124.46438, P2T_Suction := 34.86673, Superheat := 31.533272, P2T_Liquid := 59.58862, Subcool := -2.21138, Refridgerant_Type := 3);
   PCV_101_Auto_Manual : BOOL;
   PCV_101_Condenser_Pressure_PIDE : PID_ENHANCED := (PV := 163.45125, PVEUMax := 455.0, PVEUMin := -20.0, SPProg := 150.0, SPOper := 163.45125, SPHLimit := 455.0, SPLLimit := -20.0, RatioProg := 1.0, RatioOper := 1.0, RatioHLimit := 1.0, RatioLLimit := 1.0, CVEUMax := 20000.0, CVEUMin := 4000.0, CVHLimit := 100.0, HandFB := 100.0, ControlAction := 1, PGain := 4.0, IGain := 40.0, PVEDerivative := 1, PVTracking := 1, ProgOverrideReq := 1, RTSTime := 1, CVEU := 4000.0, SP := 163.45125, SPPercent := 38.621315, PVPercent := 38.621315, InitPrimary := 1, Ratio := 1.0, ProgOper := 1, Override := 1, DeltaT := 0.5);
   PCV_101_Flush_Limit : REAL := 70.0;   // Temperature Limit (Deg F) to force Condenser Water Flush
   PCV_101_Flush_Position : REAL := 20000.0;   // PCV-101 Desired Flush Position (4000-20000 counts)
   PCV_101_Flush_Time_Remaining : DINT := 30;
   PCV_101_Flush_Timer : TIMER := (PRE := 30000);   // PCV-101 Condenser Hot Water Flush Timer
   PCV_101_go_to_start_position : BOOL;
   PCV_101_Manual_Output : REAL := 100.0;
   PCV_101_Multiplexer : DINT := 1;   // Selects controlling input to multiplxer
   PCV_101_Pressure_SP : REAL := 150.0;
   PCV_101_Run_PIDE : BOOL;
   PCV_101_Start_Position : REAL := 12000.0;   // PCV-101 Desired Start Position (4000-20000 counts)
   PCV_101_Stop_PIDE : BOOL := 1;
   PLC_DateTime : DINT[7] := ([0] := 2026, [1] := 8, [2] := 24, [3] := 17, [4] := 17, [5] := 26, [6] := 851406);
        [0]   // year
        [1]   // month
        [2]   // day
        [3]   // hour
        [4]   // minute
        [5]   // seconds
        [6]   // microseconds
   PM_101 : ALIAS FOR Local:1:I.Data.1;
   PM_101_StartupTMR : TIMER := (PRE := 30000, ACC := 30002, EN := 1, DN := 1);   // PM-101 Phase Monitor Startup Delay Alarm Timer
   Process_Pump_Diff_Pressure : REAL := -3.960312;
   PT_101 : BL_Analog_Input := (Scale_20mA := 145.0, Output := 24.930937, Fault_Delay := 5);   // Process Supply Pressure
   PT_102 : BL_Analog_Input := (Scale_4mA := -7.3, Scale_20mA := 101.5, Output := 110.7004);   // R404A Compressor Suction Pressure
   PT_102_PID_Scale_Max : REAL := 121.5;
   PT_102_PID_Scale_Min : REAL := -27.3;
   PT_103 : BL_Analog_Input := (Scale_20mA := 435.0, Output := 163.45125, Fault_Delay := 5);   // R404A Compressor Discharge Pressure
   PT_103_PID_Scale_Max : REAL := 455.0;
   PT_103_PID_Scale_Min : REAL := -20.0;
   PT_104 : BL_Analog_Input := (Scale_4mA := -7.3, Scale_20mA := 101.5, Output := 110.693596);   // R404A Evaporator Suction Pressure
   PT_104_PID_Scale_Max : REAL := 121.5;
   PT_104_PID_Scale_Min : REAL := -27.3;
   PT_105 : BL_Analog_Input := (Scale_20mA := 145.0, Output := 28.855);   // Condenser Chilled Glycol Return Pressure
   PT_106 : BL_Analog_Input := (Scale_20mA := 145.0, Output := 47.868122);   // Condenser Chilled Glycol Supply Pressure
   PT_107 : BL_Analog_Input := (Scale_20mA := 145.0, Output := 25.1575);   // Process Pump Suction Pressure
   PT_108 : BL_Analog_Input := (Scale_20mA := 145.0, Output := 24.813124);   // Process Pump Suction Discharge Pressure
   Pump_1_Low_Press_Delay : TIMER := (PRE := 30000);
   Pump_High_Pressure_Alarm_Setpoint : REAL := 120.0;
   Pump_Low_Pressure_Alarm_Setpoint : REAL := 10.0;
   Pump_Manual_Release : BOOL := 1;
   Pump_Manual_Release_Timer : TIMER := (PRE := 5000, ACC := 5001, EN := 1, DN := 1);
   Pump_OK_To_Run : BOOL := 1;
   Pump_RP_ALM_TMR : TIMER := (PRE := 3000);
   Pump_Running : BOOL;
   Purge_Request : BOOL;   // Oil Management, Request to Purge
   R404A_HG_Switch_Delay : TIMER := (PRE := 10000);
   R404A_HG_Switch_Off_Delay : TIMER := (PRE := 10000);
   R404A_High_Pressure_Setpoint : REAL := 350.0;
   R404A_High_SH_Setpoint : REAL := 80.0;
   R404A_High_Superheat_Timer : TIMER := (PRE := 120000);
   R404A_Hot_Gas_Toggle : BOOL;
   R404A_Hot_Gas_Toggle_Req : BOOL;
   R404A_Low_Pressure_Delay : TIMER := (PRE := 120000);
   R404A_Low_Pressure_Setpoint : REAL := 15.0;
   R404A_Low_SC_Setpoint : REAL;
   R404A_Low_SH_Setpoint : REAL := 2.0;
   R404A_Low_Subcooling_Timer : TIMER := (PRE := 120000);
   R404A_Low_Superheat_Timer : TIMER := (PRE := 120000);
   R404A_Oil_Purge_Retires_Enable : BOOL;   // Oil Management, Oil Purge Retries Enabled
   R404A_OK_To_Run : BOOL;
   R404A_One_Comp_Running : BOOL;
   R404A_TCV_Toggle_SP_OFF : REAL := 58.0;
   R404A_TCV_Toggle_SP_ON : REAL := 62.0;
   R404A_TCV_Valve_Toggle : BOOL;
   Ramp_Soak_Current_HMI : DINT := 2#0000_0000_0000_0000_0000_0000_0000_0001;
   Ramp_Soak_Segments_HMI : DINT := 2#0000_0000_0000_0000_0000_0000_0011_1110;
   Ramp_Soak_Segments_HMI_Set : REAL := 5.0;
   REACTOR_BATCH_PID_START : BOOL;
   REACTOR_BATCH_PID_STOP : BOOL := 1;
   REACTOR_BATCH_PIDE : PID_ENHANCED := (PV := 20.0, PVEUMax := 200.0, PVEUMin := -40.0, SPProg := 20.0, SPOper := 20.0, SPHLimit := 200.0, SPLLimit := -40.0, RatioProg := 1.0, RatioOper := 1.0, RatioHLimit := 1.0, RatioLLimit := 1.0, CVInitReq := 1, CVInitValue := 23.3, CVOper := 51.454544, CVEUMax := 50.0, CVEUMin := -5.0, CVHLimit := 100.0, PGain := 12.0, IGain := 4.0, PVEDerivative := 1, DSmoothing := 1, PVTracking := 1, AllowCasRat := 1, ProgOverrideReq := 1, RTSTime := 1, CVEU := 23.3, CV := 51.454544, CVInitializing := 1, SP := 20.0, SPPercent := 25.0, PVPercent := 25.0, InitPrimary := 1, Ratio := 1.0, Override := 1, DeltaT := 1.0);
   REACTOR_BATCH_PIDE_CV_AS_SP : REAL := 23.3;
   REACTOR_BATCH_PV : REAL := 20.0;
   REACTOR_BATCH_SP_HIGH : REAL := 50.0;
   REACTOR_BATCH_SP_LOW : REAL := -10.0;
   REACTOR_HEAT_RUN_PIDE : BOOL;
   REACTOR_HEAT_STOP_PIDE : BOOL := 1;
   REACTOR_HEATERS_OK_TO_RUN : BOOL;
   REACTOR_HEATERS_TEMPERATURE_PIDE : PID_ENHANCED := (PV := 23.3, PVEUMax := 200.0, PVEUMin := -40.0, SPProg := 20.0, SPOper := 23.3, SPCascade := 23.3, SPHLimit := 200.0, SPLLimit := -40.0, RatioProg := 1.0, RatioOper := 1.0, RatioHLimit := 1.0, RatioLLimit := 1.0, CVEUMax := 20000.0, CVEUMin := 4000.0, CVHLimit := 100.0, HandFB := 78.0, PGain := 12.0, IGain := 3.0, PVEDerivative := 1, PVTracking := 1, AllowCasRat := 1, ProgOverrideReq := 1, RTSTime := 1, CVEU := 4000.0, SP := 23.3, SPPercent := 26.374998, PVPercent := 26.374998, InitPrimary := 1, Ratio := 1.0, ProgOper := 1, Override := 1, DeltaT := 1.0);
   Regulate_Request : BOOL;
   Remote_Alarm_Reset : BOOL;
   Remote_Enable_Batch : BOOL;   // Remote Jacket/Batch Control (0=Jacket, 1=Batch)
   Remote_Enable_Batchx : DINT;   // Remote Jacket/Batch Control (0=Jacket, 1=Batch)
   Remote_System_Start : BOOL;   // Remote Start/Stop 0=Stop 1=Start
   Remote_Temp_Setpoint : REAL := 25.0;   // Remote Temperature Setpoint
   RX_Profile_Stop_SP_Control : TIMER := (PRE := 5000, ACC := 5002, EN := 1, DN := 1);
   RX_RMPS : RAMP_SOAK := (PV := 23.3, NumberOfSegs := 6, TimeRate := 1, RampDeadband := 1.0, SoakDeadband := 1.0, OutProg := 20.0, OutOper := 20.0, ProgManualReq := 1, Out := 20.0, ProgOper := 1, Manual := 1);
   RX_RMPS_Current_Segment : DINT;
   RX_RMPS_Output : REAL := 20.0;
   RX_RMPS_Ramp_Value : REAL[11] := ([1] := 2.0, [2] := 2.0, [3] := 2.0, [4] := 2.0, [5] := 2.0);
   RX_RMPS_Soak_Time : REAL[11] := ([1] := 2.0, [2] := 2.0, [3] := 2.0, [4] := 2.0, [5] := 2.0);
   RX_RMPS_Soak_Value : REAL[11] := ([0] := 23.3, [2] := 5.0, [3] := 10.0, [4] := 15.0, [5] := 20.0);
   RX_RMPS_SP_Out : REAL := 20.0;
   RX_Run_Temp_Profile : BOOL;
   RX_Start_Temperature_Profile : BOOL;
   RX_Stop_Temp_Profile : BOOL := 1;
   SCR_101_Auto_Manual : BOOL;
   SCR_101_Manual_Output : REAL := 78.0;
   SCR_Output_Percent : DINT;
   SCR_PID_Request : REAL;
   Sensor_1 : BudLib_Analog_Sensor := (Raw_Data := 6751.0, Fault_Disable := 1);
   Sensor_10 : BudLib_Analog_Sensor := (Raw_Data := 5038.0, Fault_Disable := 1);
   Sensor_2 : BudLib_Analog_Sensor := (Raw_Data := 21353.0, Disable_High_Fault := 1, Fault_Disable := 1);
   Sensor_3 : BudLib_Analog_Sensor := (Raw_Data := 10012.0, Fault_Disable := 1);
   Sensor_4 : BudLib_Analog_Sensor := (Raw_Data := 21352.0, Disable_High_Fault := 1, Fault_Disable := 1);
   Sensor_5 : BudLib_Analog_Sensor := (Raw_Data := 7181.0, Disable_High_Fault := 1, Fault_Disable := 1);
   Sensor_6 : BudLib_Analog_Sensor := (Raw_Data := 9292.0, Disable_High_Fault := 1, Fault_Disable := 1);
   Sensor_7 : BudLib_Analog_Sensor := (Raw_Data := 6776.0, Fault_Disable := 1);
   Sensor_8 : BudLib_Analog_Sensor := (Raw_Data := 6738.0, Fault_Disable := 1);
   Sensor_9 : BudLib_Analog_Sensor := (Raw_Data := 4018.0, Disable_High_Fault := 1, Fault_Disable := 1);
   Short_Cycle_1_Time_Remaining : DINT;
   Short_Cycle_2_Time_Remaining : DINT;
   Short_Cycle_3_Time_Remaining : DINT;
   Short_Cycle_Timer_1 : TIMER := (PRE := 180000, ACC := 2207);
   Slot_2_Status : DINT := 16384;
   Slot_3_Status : DINT := 16384;
   Slot_4_Status : DINT := 16384;
   Slot_5_Status : DINT := 16384;
   Slot_6_Status : DINT := 16384;
   Slot_7_Status : DINT := 16384;
   Slot_8_Status : DINT := 16384;
   Slot_9_Status : DINT := 16384;
   Start_Up_Delay : TIMER := (PRE := 15000, ACC := 15002, EN := 1, DN := 1);
   System_Mode : BOOL;   // 0 = Local Control 1 = Remote Control
   System_Start : BOOL;   // System Start
   T_SENSOR_1 : BudLib_Analog_Sensor := (Raw_Data := 233.0, Sensor_Type := 1, Fault_Disable := 1);
   T_SENSOR_10 : BudLib_Analog_Sensor := (Raw_Data := 8700.0, Sensor_Type := 1, Sensor_Alarm := 1, Fault_Disable := 1);
   T_SENSOR_2 : BudLib_Analog_Sensor := (Raw_Data := 221.0, Sensor_Type := 1, Fault_Disable := 1);
   T_SENSOR_3 : BudLib_Analog_Sensor := (Raw_Data := 737.0, Sensor_Type := 1, Fault_Disable := 1);
   T_SENSOR_4 : BudLib_Analog_Sensor := (Raw_Data := 751.0, Sensor_Type := 1, Fault_Disable := 1);
   T_SENSOR_5 : BudLib_Analog_Sensor := (Raw_Data := 851.0, Sensor_Type := 1, Fault_Disable := 1);
   T_SENSOR_6 : BudLib_Analog_Sensor := (Raw_Data := 734.0, Sensor_Type := 1, Fault_Disable := 1);
   T_SENSOR_7 : BudLib_Analog_Sensor := (Raw_Data := -149.0, Sensor_Type := 1, Fault_Disable := 1);
   T_SENSOR_8 : BudLib_Analog_Sensor := (Raw_Data := 715.0, Sensor_Type := 1, Fault_Disable := 1);
   T_SENSOR_9 : BudLib_Analog_Sensor := (Raw_Data := 688.0, Sensor_Type := 1);
   TCM_FROM_DCS : DINT[4] := ([1] := 210, [2] := 20);   // Data from TCU to Supervisory System
        [0]   // Control Bits from Supervisory System ModBus 40010
        [0].0   // Heartbeat Return
        [0].1   // Remote Start/Stop
        [0].2   // Remote Jacket/Batch Control
        [0].3   // Remote Alarm Reset
        [1]   // Remote Temperature Setpoint
        [2]   // Spare
   TCM_TO_DCS : DINT[10] := ([1] := 198, [2] := 202, [3] := 190, [4] := 10, [5] := 219);   // Data to TCU from Supervisory System
        [0]   // NOT USED
        [0].0   // Heartbeat
        [0].1   // Local/Remote Status 0 = Local Control 1 = Remote Control
        [0].2   // Batch/Jacket Mode 0=Jacket 1=Batch
        [0].3   // Process Pump Running
        [0].4   // TCM Heating
        [0].5   // TCM Cooling
        [0].6   // Alarms Present
        [0].7   // spare
        [0].8   // spare
        [1]   // TCM Outlet Temperature TE-101 (0.1 Scale)
        [2]   // TCP Return Pressure TE-102 (0.1 Scale)
        [3]   // Process Supply Pressure PT-101 (0.1 Scale)
        [4]   // Active Temperature Setpoint (0.1 Scale)
        [5]   // Vessel Temperature (0.1 Scale)
        [6]   // Spare
        [7]   // Spare
        [8]   // Spare
   TCV_101_Auto_Manual : BOOL;
   TCV_101_CV_RAW : ALIAS FOR Local:7:O.Ch3Data;   // TCV-101 Valve De-Scale Output (4000-20000)
   TCV_101_EVAP_PRESSURE_PIDE : PID_ENHANCED := (PV := 110.693596, PVEUMax := 122.0, PVEUMin := -27.0, SPProg := 25.0, SPOper := 101.5, SPHLimit := 101.5, SPLLimit := -7.3, RatioProg := 1.0, RatioOper := 1.0, RatioHLimit := 1.0, RatioLLimit := 1.0, CVEUMax := 20000.0, CVEUMin := 4000.0, CVHLimit := 100.0, CVLLimit := 8.0, HandFB := 8.0, PGain := 2.0, IGain := 10.0, PVEDerivative := 1, DSmoothing := 1, PVTracking := 1, AllowCasRat := 1, ProgCasRatReq := 1, ProgOverrideReq := 1, RTSTime := 1, CVEU := 4000.0, CVLAlarm := 1, SP := 101.5, SPPercent := 86.24161, SPHAlarm := 1, PVPercent := 92.41182, E := -9.193596, EPercent := -6.170212, InitPrimary := 1, WindupHOut := 1, WindupLOut := 1, Ratio := 1.0, ProgOper := 1, Override := 1, DeltaT := 1.0);   // TCV-101 Hot Gas Pressure PID loop
   TCV_101_EVAP_TEMPERATURE_PIDE : PID_ENHANCED := (PV := 23.3, PVEUMax := 200.0, PVEUMin := -40.0, SPProg := 20.0, SPOper := 23.3, SPCascade := 23.3, SPHLimit := 200.0, SPLLimit := -40.0, RatioProg := 1.0, RatioOper := 1.0, RatioHLimit := 1.0, RatioLLimit := 1.0, CVEUMax := 20000.0, CVEUMin := 4000.0, CVHLimit := 100.0, CVLLimit := 8.0, HandFB := 8.0, PGain := 50.0, IGain := 20.0, PVEDerivative := 1, DSmoothing := 1, PVTracking := 1, AllowCasRat := 1, ProgOverrideReq := 1, RTSTime := 1, CVEU := 4000.0, CVLAlarm := 1, SP := 23.3, SPPercent := 26.374998, PVPercent := 26.374998, InitPrimary := 1, WindupLOut := 1, Ratio := 1.0, ProgOper := 1, Override := 1, DeltaT := 1.0);   // TCV-101 Evaporator Hot Gas Bypass PID loop
   TCV_101_High_Range_CV_Max : REAL := 100.0;
   TCV_101_High_Range_CV_Min : REAL := 8.0;
   TCV_101_Low_Range_CV_Max : REAL := 100.0;
   TCV_101_Low_Range_CV_Min : REAL := 5.0;
   TCV_101_Manual_Output : REAL := 8.0;
   TCV_101_Mid_Range_CV_Max : REAL := 100.0;
   TCV_101_Mid_Range_CV_Min : REAL := 8.0;
   TCV_101_Output_Percent : REAL;
   TCV_101_Pressure_Setpoint : REAL := 25.0;   // TCV-101 Hot Gas Pressure PID loop Setpoint
   TCV_101_Relay : BOOL;
   TCV_101_Run_PIDE : BOOL;
   TCV_101_Stop_PIDE : BOOL := 1;
   TCV_102_CV_RAW : ALIAS FOR Local:8:O.Ch0Data;   // TCV-102 Valve De-Scale Output (4000-20000)
   TCV_102_Relay : BOOL;
   TCV_CV : REAL;   // TCV Loop Output Scaled (0-100%)
   TCV_Multiplexer : DINT := 1;
   TCV_Mux : MULTIPLEXER := (In1 := 4000.0, In2 := 4000.0, In3 := 8800.0, Selector := 1, Out := 4000.0);
   TE_101 : BL_Analog_Input := (Output := 23.3);   // Process Supply Temperature
   TE_101_PID_Scale_Max : REAL := 20.0;
   TE_101_PID_Scale_Min : REAL := -20.0;
   TE_102 : BL_Analog_Input := (Output := 22.1);   // Process Return Temperature
   TE_103 : BL_Analog_Input := (Output := 73.7);   // R507A Liquid Line Temperature
   TE_104 : BL_Analog_Input := (Output := 75.1);   // R507A Evaporator Suction Temperature
   TE_105 : BL_Analog_Input := (Output := 85.1);   // R507A Compressor Suction Temperature
   TE_106 : BL_Analog_Input := (Output := 73.4);   // CONDENSER CHILLED GLYCOL OUTLET TEMPERATURE SENSOR
   TE_108 : BL_Analog_Input := (Output := 71.5);   // CONDENSER CHILLED GLYCOL INLET TEMPERATURE SENSOR
   Temperature_Setpoint : REAL := 20.0;
   Temperature_Setpoint_Last : REAL := 20.0;
   Temperature_Setpoint_Max : REAL := 85.0;   // Maximum Operating Temperature Setpoint (Deg C)
   Temperature_Setpoint_Min : REAL := -5.0;   // Minimum Operating Temperature Setpoint (Deg C)
   test_th : DINT;
   TSH_101 : ALIAS FOR Local:1:I.Data.4;
   Valve_delay_count : REAL;
   Valve_Flush_SP : REAL := 13600.0;
   VESSEL_TEMPERATURE : BL_Analog_Input := (Scale_4mA := -50.0, Scale_20mA := 200.0, Output := 20.0, Fault_Delay := 5);   // End User Reactor Temperature
END_VAR

PROGRAM A_MainProgram   (* main routine Routine_Schedule *)

ROUTINE Alarms_Setup   (* ladder *)
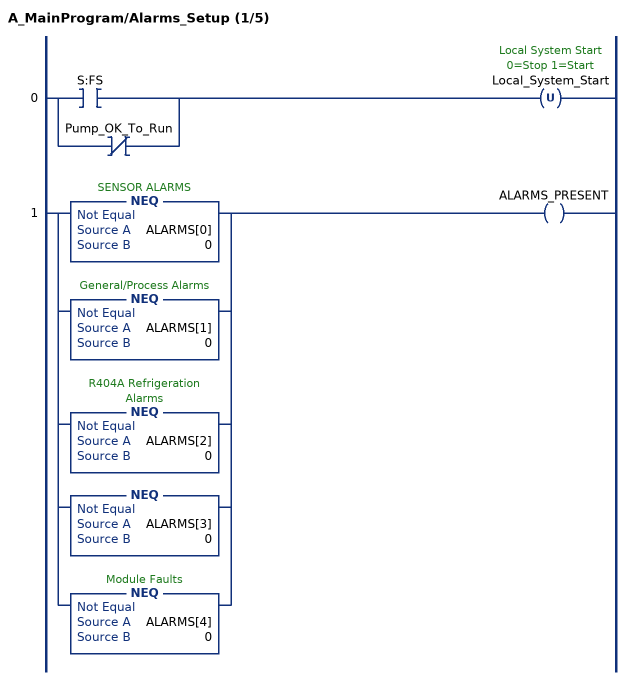
   0: [XIC(S:FS) ,XIO(Pump_OK_To_Run) ]OTU(Local_System_Start);
   1: [NEQ(ALARMS[0],0) ,NEQ(ALARMS[1],0) ,NEQ(ALARMS[2],0) ,NEQ(ALARMS[3],0) ,NEQ(ALARMS[4],0) ]OTE(ALARMS_PRESENT);
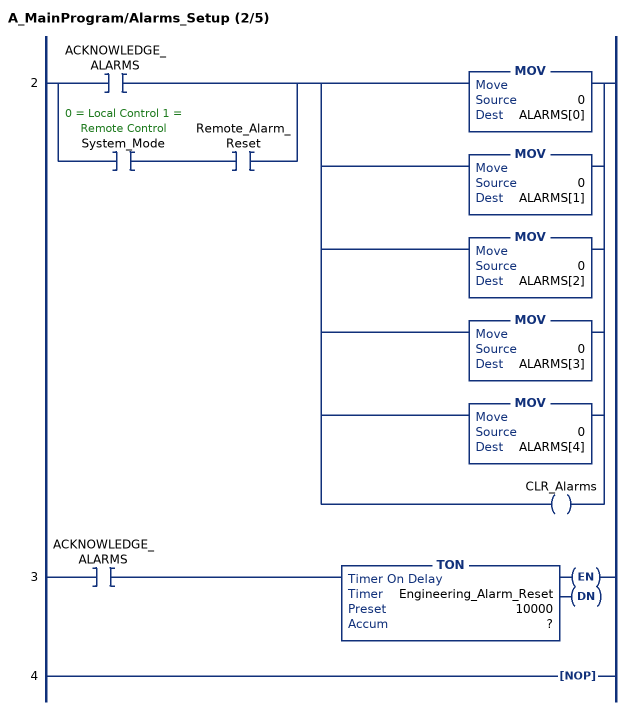
   2: [XIC(ACKNOWLEDGE_ALARMS) ,XIC(System_Mode) XIC(Remote_Alarm_Reset) ][MOV(0,ALARMS[0]) ,MOV(0,ALARMS[1]) ,MOV(0,ALARMS[2]) ,MOV(0,ALARMS[3]) ,MOV(0,ALARMS[4]) ,OTE(CLR_Alarms) ];
   3: XIC(ACKNOWLEDGE_ALARMS)TON(Engineering_Alarm_Reset,?,?);
   4: NOP();
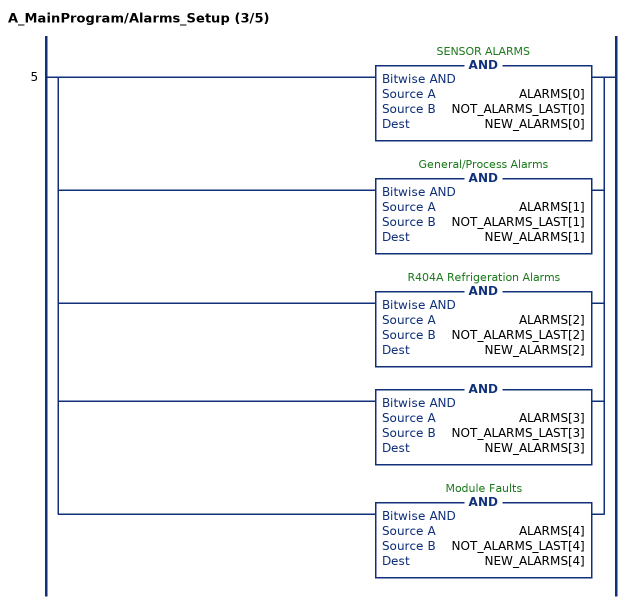
   5: [AND(ALARMS[0],NOT_ALARMS_LAST[0],NEW_ALARMS[0]) ,AND(ALARMS[1],NOT_ALARMS_LAST[1],NEW_ALARMS[1]) ,AND(ALARMS[2],NOT_ALARMS_LAST[2],NEW_ALARMS[2]) ,AND(ALARMS[3],NOT_ALARMS_LAST[3],NEW_ALARMS[3]) ,AND(ALARMS[4],NOT_ALARMS_LAST[4],NEW_ALARMS[4]) ];
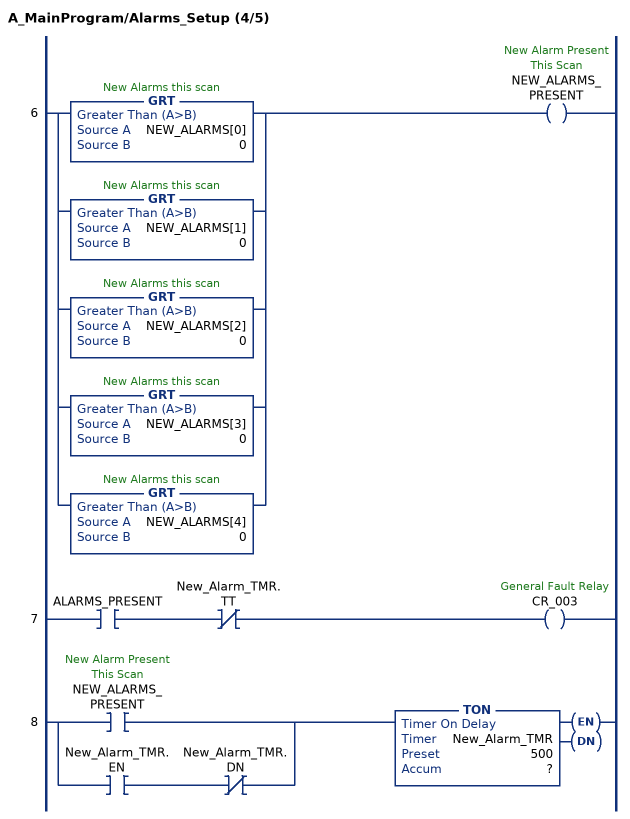
   6: [GRT(NEW_ALARMS[0],0) ,GRT(NEW_ALARMS[1],0) ,GRT(NEW_ALARMS[2],0) ,GRT(NEW_ALARMS[3],0) ,GRT(NEW_ALARMS[4],0) ]OTE(NEW_ALARMS_PRESENT);
   7: XIC(ALARMS_PRESENT)XIO(New_Alarm_TMR.TT)OTE(CR_003);
   8: [XIC(NEW_ALARMS_PRESENT) ,XIC(New_Alarm_TMR.EN) XIO(New_Alarm_TMR.DN) ]TON(New_Alarm_TMR,?,?);
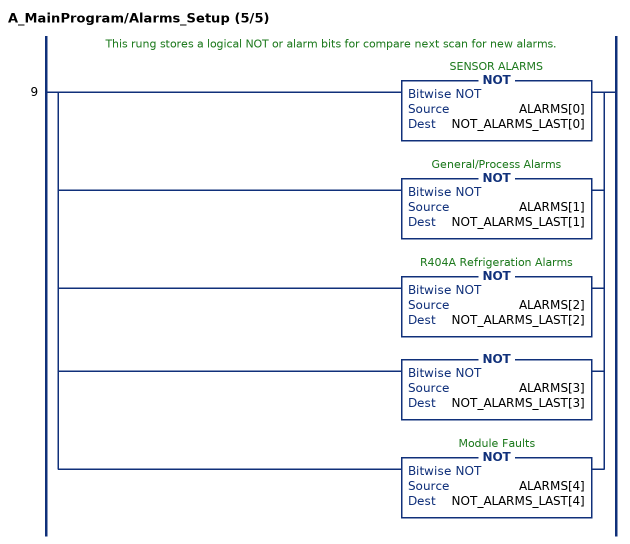
   // This rung stores a logical NOT or alarm bits for compare next scan for new alarms.
   9: [NOT(ALARMS[0],NOT_ALARMS_LAST[0]) ,NOT(ALARMS[1],NOT_ALARMS_LAST[1]) ,NOT(ALARMS[2],NOT_ALARMS_LAST[2]) ,NOT(ALARMS[3],NOT_ALARMS_LAST[3]) ,NOT(ALARMS[4],NOT_ALARMS_LAST[4]) ];
END_ROUTINE

ROUTINE DCS_COMM   (* ladder *)
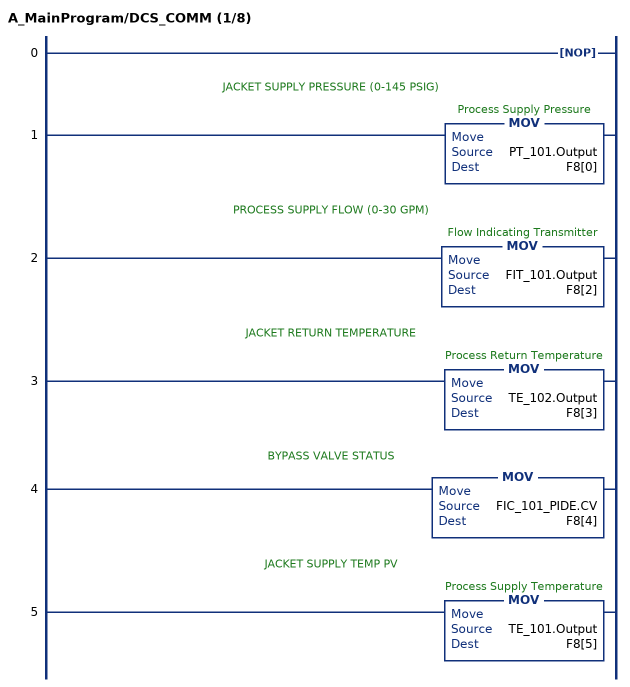
   0: NOP();
   // JACKET SUPPLY PRESSURE (0-145 PSIG)
   1: MOV(PT_101.Output,F8[0]);
   // PROCESS SUPPLY FLOW (0-30 GPM)
   2: MOV(FIT_101.Output,F8[2]);
   // JACKET RETURN TEMPERATURE
   3: MOV(TE_102.Output,F8[3]);
   // BYPASS VALVE STATUS
   4: MOV(FIC_101_PIDE.CV,F8[4]);
   // JACKET SUPPLY TEMP PV
   5: MOV(TE_101.Output,F8[5]);
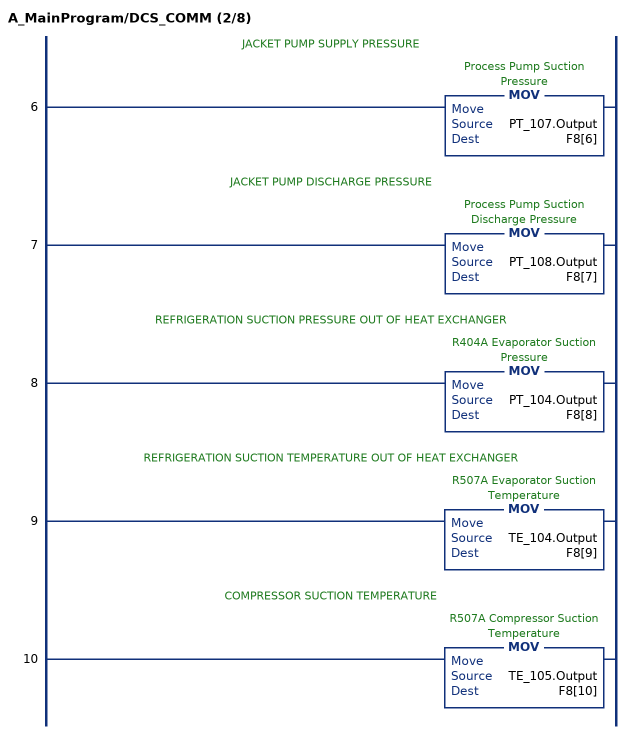
   // JACKET PUMP SUPPLY PRESSURE
   6: MOV(PT_107.Output,F8[6]);
   // JACKET PUMP DISCHARGE PRESSURE
   7: MOV(PT_108.Output,F8[7]);
   // REFRIGERATION SUCTION PRESSURE OUT OF HEAT EXCHANGER
   8: MOV(PT_104.Output,F8[8]);
   // REFRIGERATION SUCTION TEMPERATURE OUT OF HEAT EXCHANGER
   9: MOV(TE_104.Output,F8[9]);
   // COMPRESSOR SUCTION TEMPERATURE
   10: MOV(TE_105.Output,F8[10]);
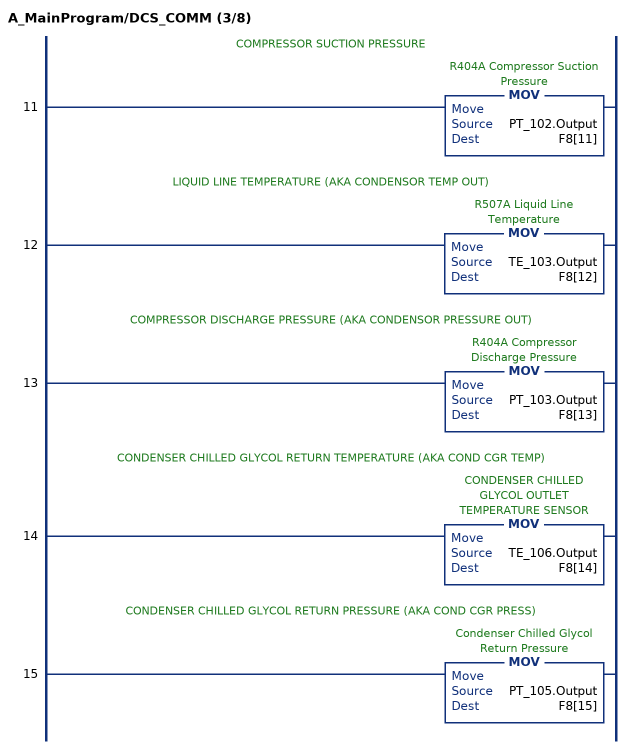
   // COMPRESSOR SUCTION PRESSURE
   11: MOV(PT_102.Output,F8[11]);
   // LIQUID LINE TEMPERATURE (AKA CONDENSOR TEMP OUT)
   12: MOV(TE_103.Output,F8[12]);
   // COMPRESSOR DISCHARGE PRESSURE (AKA CONDENSOR PRESSURE OUT)
   13: MOV(PT_103.Output,F8[13]);
   // CONDENSER CHILLED GLYCOL RETURN TEMPERATURE (AKA COND CGR TEMP)
   14: MOV(TE_106.Output,F8[14]);
   // CONDENSER CHILLED GLYCOL RETURN PRESSURE (AKA COND CGR PRESS)
   15: MOV(PT_105.Output,F8[15]);
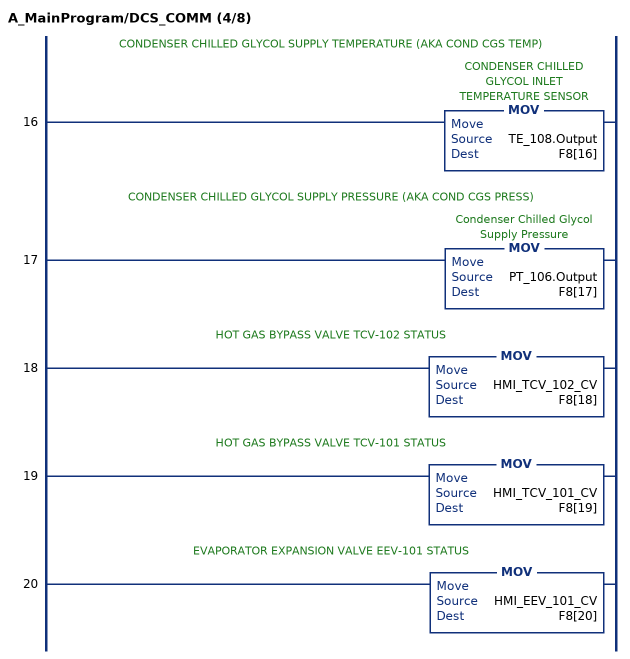
   // CONDENSER CHILLED GLYCOL SUPPLY TEMPERATURE (AKA COND CGS TEMP)
   16: MOV(TE_108.Output,F8[16]);
   // CONDENSER CHILLED GLYCOL SUPPLY PRESSURE (AKA COND CGS PRESS)
   17: MOV(PT_106.Output,F8[17]);
   // HOT GAS BYPASS VALVE TCV-102 STATUS
   18: MOV(HMI_TCV_102_CV,F8[18]);
   // HOT GAS BYPASS VALVE TCV-101 STATUS
   19: MOV(HMI_TCV_101_CV,F8[19]);
   // EVAPORATOR EXPANSION VALVE EEV-101 STATUS
   20: MOV(HMI_EEV_101_CV,F8[20]);
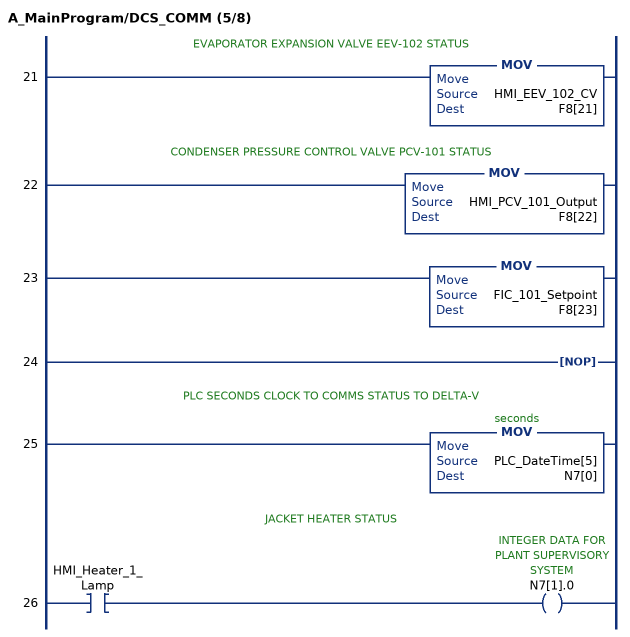
   // EVAPORATOR EXPANSION VALVE EEV-102 STATUS
   21: MOV(HMI_EEV_102_CV,F8[21]);
   // CONDENSER PRESSURE CONTROL VALVE PCV-101 STATUS
   22: MOV(HMI_PCV_101_Output,F8[22]);
   23: MOV(FIC_101_Setpoint,F8[23]);
   24: NOP();
   // PLC SECONDS CLOCK TO COMMS STATUS TO DELTA-V
   25: MOV(PLC_DateTime[5],N7[0]);
   // JACKET HEATER STATUS
   26: XIC(HMI_Heater_1_Lamp)OTE(N7[1].0);
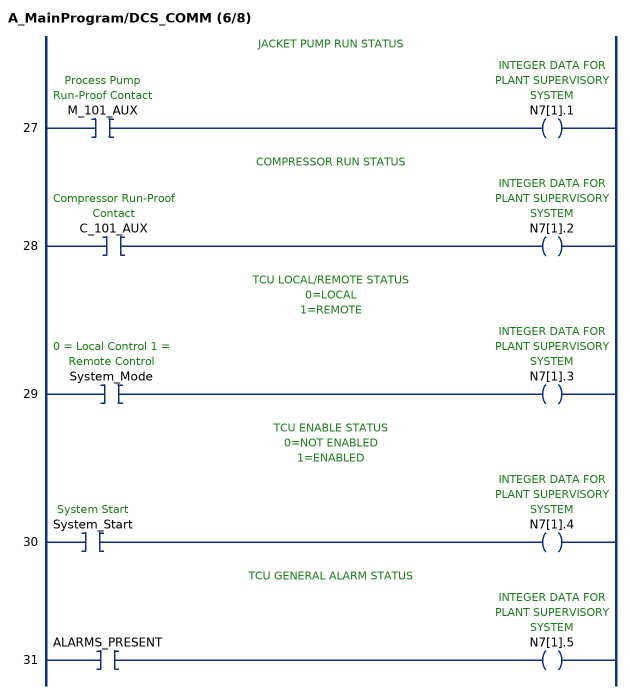
   // JACKET PUMP RUN STATUS
   27: XIC(M_101_AUX)OTE(N7[1].1);
   // COMPRESSOR RUN STATUS
   28: XIC(C_101_AUX)OTE(N7[1].2);
   // TCU LOCAL/REMOTE STATUS
   // 0=LOCAL
   // 1=REMOTE
   29: XIC(System_Mode)OTE(N7[1].3);
   // TCU ENABLE STATUS
   // 0=NOT ENABLED
   // 1=ENABLED
   30: XIC(System_Start)OTE(N7[1].4);
   // TCU GENERAL ALARM STATUS
   31: XIC(ALARMS_PRESENT)OTE(N7[1].5);
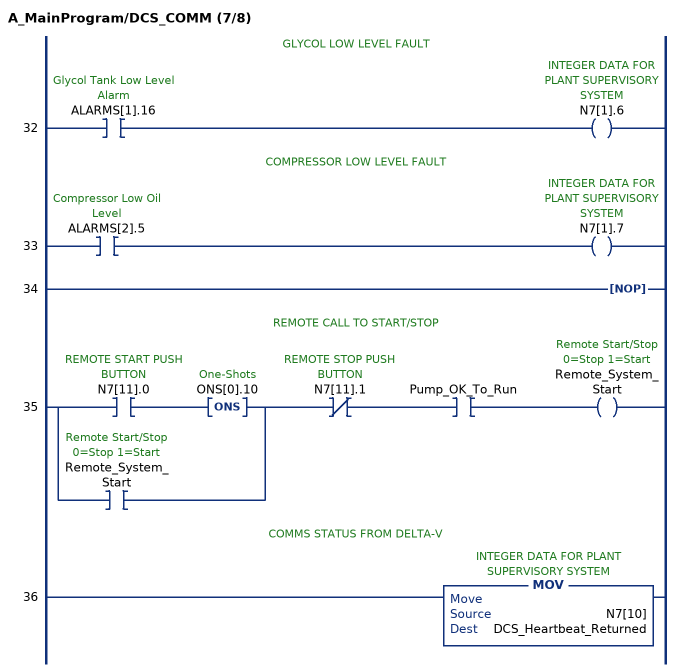
   // GLYCOL LOW LEVEL FAULT
   32: XIC(ALARMS[1].16)OTE(N7[1].6);
   // COMPRESSOR LOW LEVEL FAULT
   33: XIC(ALARMS[2].5)OTE(N7[1].7);
   34: NOP();
   // REMOTE CALL TO START/STOP
   35: [XIC(N7[11].0) ONS(ONS[0].10) ,XIC(Remote_System_Start) ]XIO(N7[11].1)XIC(Pump_OK_To_Run)OTE(Remote_System_Start);
   // COMMS STATUS FROM DELTA-V
   36: MOV(N7[10],DCS_Heartbeat_Returned);
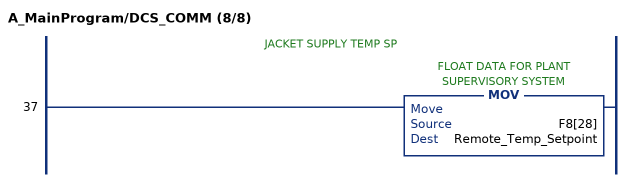
   // JACKET SUPPLY TEMP SP
   37: MOV(F8[28],Remote_Temp_Setpoint);
END_ROUTINE
